(* IEC 61131-3 sources: plc-st-coding-agent/progress/evidence/f14_v10_full_20261113/jobs/custom_deepseek-v4pro (part 4) *)

(* ---- public-medium-02.raw_candidate_01.st ---- *)
TYPE ST_AnalogChannel :
STRUCT
    enable : BOOL;
    hiLIM : REAL;
    loLIM : REAL;
    bipolar : BOOL;
    measuringMode : INT;
    retVal : WORD;
    outputValue : REAL;
END_STRUCT
END_TYPE

(*
ENGINEERING_CONTRACT
Activation: process first count ordinal channels, count >= 0, clamped to min array lengths.
Enable: only channels[].enable = TRUE is evaluated; disabled rows retain previous retVal/outputValue.
retVal: for enabled rows write WORD#0 on success; WORD#16#8001 invalid measuringMode (PUB006); WORD#16#8002 hiLIM<=loLIM (PUB007).
Priority/simultaneous checks: measuringMode validity checked before hiLIM<=loLIM; simultaneous invalid mode and bad limits yields 16#8001 (unspecified, chosen).
outputValue: written only for enabled successful conversions; mode0 linear scaling clamped to 0/27648 or -27648/27648 (PUB003); mode1 raw/10 (PUB004); mode2 raw/100 (PUB005).
Read-only: analogValues unchanged; configuration fields only read (PUB001, PUB002).
Bounds: match by ordinal from each array lower bound; invalid count processes none.
Units: raw INT, output REAL, limits REAL; no time.
*)

(* CONTRACT_RULES [] *)

FUNCTION_BLOCK AnalogBatchProcessing
VAR_INPUT
    count : DINT;
END_VAR
VAR_IN_OUT
    analogValues : ARRAY[*] OF INT;
    channels : ARRAY[*] OF ST_AnalogChannel;
END_VAR
VAR
    tmp_lbA : DINT;
    tmp_lbC : DINT;
    tmp_availA : DINT;
    tmp_availC : DINT;
    tmp_process : DINT;
    tmp_i : DINT;
    tmp_idxA : DINT;
    tmp_idxC : DINT;
    tmp_raw : INT;
    tmp_rawReal : REAL;
    tmp_frac : REAL;
END_VAR

tmp_lbA := LOWER_BOUND(analogValues, 1);
tmp_lbC := LOWER_BOUND(channels, 1);
tmp_availA := UPPER_BOUND(analogValues, 1) - tmp_lbA + 1;
tmp_availC := UPPER_BOUND(channels, 1) - tmp_lbC + 1;

tmp_process := count;
IF tmp_process < 0 THEN
    tmp_process := 0;
END_IF;
IF tmp_process > tmp_availA THEN
    tmp_process := tmp_availA;
END_IF;
IF tmp_process > tmp_availC THEN
    tmp_process := tmp_availC;
END_IF;

FOR tmp_i := 0 TO tmp_process - 1 DO
    tmp_idxA := tmp_lbA + tmp_i;
    tmp_idxC := tmp_lbC + tmp_i;

    IF channels[tmp_idxC].enable THEN
        channels[tmp_idxC].retVal := WORD#0;

        IF (channels[tmp_idxC].measuringMode < 0) OR (channels[tmp_idxC].measuringMode > 2) THEN
            channels[tmp_idxC].retVal := WORD#16#8001;
            (* skip conversion; outputValue unchanged *)
        ELSIF channels[tmp_idxC].hiLIM <= channels[tmp_idxC].loLIM THEN
            channels[tmp_idxC].retVal := WORD#16#8002;
            (* skip conversion; outputValue unchanged *)
        ELSE
            tmp_raw := analogValues[tmp_idxA];
            tmp_rawReal := INT_TO_REAL(tmp_raw);

            CASE channels[tmp_idxC].measuringMode OF
                0:
                    IF channels[tmp_idxC].bipolar THEN
                        IF tmp_rawReal < -27648.0 THEN
                            tmp_rawReal := -27648.0;
                        ELSIF tmp_rawReal > 27648.0 THEN
                            tmp_rawReal := 27648.0;
                        END_IF;
                        tmp_frac := (tmp_rawReal + 27648.0) / 55296.0;
                    ELSE
                        IF tmp_rawReal < 0.0 THEN
                            tmp_rawReal := 0.0;
                        ELSIF tmp_rawReal > 27648.0 THEN
                            tmp_rawReal := 27648.0;
                        END_IF;
                        tmp_frac := tmp_rawReal / 27648.0;
                    END_IF;

                    channels[tmp_idxC].outputValue := channels[tmp_idxC].loLIM
                        + tmp_frac * (channels[tmp_idxC].hiLIM - channels[tmp_idxC].loLIM);

                1:
                    channels[tmp_idxC].outputValue := tmp_rawReal / 10.0;

                2:
                    channels[tmp_idxC].outputValue := tmp_rawReal / 100.0;

                ELSE
                    (* unreachable due to mode check above *)
                END_CASE;
        END_IF;
    END_IF;
END_FOR;

END_FUNCTION_BLOCK

(* ---- public-medium-02.raw_candidate_02.st ---- *)
TYPE ST_AnalogChannel :
STRUCT
    enable : BOOL;
    hiLIM : REAL;
    loLIM : REAL;
    bipolar : BOOL;
    measuringMode : INT;
    retVal : WORD;
    outputValue : REAL;
END_STRUCT
END_TYPE;

(*
ENGINEERING_CONTRACT
Activation: process first count ordinal channels, count >= 0, clamped to min array lengths.
Enable: only channels[].enable = TRUE is evaluated; disabled rows retain previous retVal/outputValue.
retVal: for enabled rows write WORD#0 on success; WORD#16#8001 invalid measuringMode (PUB006); WORD#16#8002 hiLIM<=loLIM (PUB007).
Priority/simultaneous checks: measuringMode validity checked before hiLIM<=loLIM; simultaneous invalid mode and bad limits yields 16#8001 (unspecified, chosen).
outputValue: written only for enabled successful conversions; mode0 linear scaling clamped to 0/27648 or -27648/27648 (PUB003); mode1 raw/10 (PUB004); mode2 raw/100 (PUB005).
Read-only: analogValues unchanged; configuration fields only read (PUB001, PUB002).
Bounds: match by ordinal from each array lower bound; invalid count processes none.
Units: raw INT, output REAL, limits REAL; no time.
*)

(* CONTRACT_RULES [] *)

FUNCTION_BLOCK AnalogBatchProcessing
VAR_INPUT
    count : DINT;
END_VAR
VAR_IN_OUT
    analogValues : ARRAY[*] OF INT;
    channels : ARRAY[*] OF ST_AnalogChannel;
END_VAR
VAR
    tmp_lbA : DINT;
    tmp_lbC : DINT;
    tmp_availA : DINT;
    tmp_availC : DINT;
    tmp_process : DINT;
    tmp_i : DINT;
    tmp_idxA : DINT;
    tmp_idxC : DINT;
    tmp_raw : INT;
    tmp_rawReal : REAL;
    tmp_frac : REAL;
END_VAR

tmp_lbA := LOWER_BOUND(analogValues, 1);
tmp_lbC := LOWER_BOUND(channels, 1);
tmp_availA := UPPER_BOUND(analogValues, 1) - tmp_lbA + 1;
tmp_availC := UPPER_BOUND(channels, 1) - tmp_lbC + 1;

tmp_process := count;
IF tmp_process < 0 THEN
    tmp_process := 0;
END_IF;
IF tmp_process > tmp_availA THEN
    tmp_process := tmp_availA;
END_IF;
IF tmp_process > tmp_availC THEN
    tmp_process := tmp_availC;
END_IF;

FOR tmp_i := 0 TO tmp_process - 1 DO
    tmp_idxA := tmp_lbA + tmp_i;
    tmp_idxC := tmp_lbC + tmp_i;

    IF channels[tmp_idxC].enable THEN
        channels[tmp_idxC].retVal := WORD#0;

        IF (channels[tmp_idxC].measuringMode < 0) OR (channels[tmp_idxC].measuringMode > 2) THEN
            channels[tmp_idxC].retVal := WORD#16#8001;
            (* skip conversion; outputValue unchanged *)
        ELSIF channels[tmp_idxC].hiLIM <= channels[tmp_idxC].loLIM THEN
            channels[tmp_idxC].retVal := WORD#16#8002;
            (* skip conversion; outputValue unchanged *)
        ELSE
            tmp_raw := analogValues[tmp_idxA];
            tmp_rawReal := INT_TO_REAL(tmp_raw);

            CASE channels[tmp_idxC].measuringMode OF
                0:
                    IF channels[tmp_idxC].bipolar THEN
                        IF tmp_rawReal < -27648.0 THEN
                            tmp_rawReal := -27648.0;
                        ELSIF tmp_rawReal > 27648.0 THEN
                            tmp_rawReal := 27648.0;
                        END_IF;
                        tmp_frac := (tmp_rawReal + 27648.0) / 55296.0;
                    ELSE
                        IF tmp_rawReal < 0.0 THEN
                            tmp_rawReal := 0.0;
                        ELSIF tmp_rawReal > 27648.0 THEN
                            tmp_rawReal := 27648.0;
                        END_IF;
                        tmp_frac := tmp_rawReal / 27648.0;
                    END_IF;

                    channels[tmp_idxC].outputValue := channels[tmp_idxC].loLIM
                        + tmp_frac * (channels[tmp_idxC].hiLIM - channels[tmp_idxC].loLIM);

                1:
                    channels[tmp_idxC].outputValue := tmp_rawReal / 10.0;

                2:
                    channels[tmp_idxC].outputValue := tmp_rawReal / 100.0;

                ELSE
                    (* unreachable due to mode check above *)
                    tmp_raw := tmp_raw;   (* dummy statement to satisfy CASE syntax *)
                END_CASE;
        END_IF;
    END_IF;
END_FOR;

END_FUNCTION_BLOCK

(* ---- public-medium-03.candidate_01.st ---- *)
FUNCTION_BLOCK FB
VAR_INPUT
    cyclicExecution : BOOL;
    trigger : BOOL;
    value : LREAL;
    windowSize : INT;
    reset : BOOL;
END_VAR
VAR_OUTPUT
    average : LREAL;
    windowSizeReached : BOOL;
    error : BOOL;
    status : WORD;
END_VAR
VAR
    local_triggerR : R_TRIG;
    local_buffer : ARRAY[0..99] OF LREAL;
    local_count : INT := 0;
    local_head : INT := 0;
    local_tail : INT := 0;
    local_sum : LREAL := 0.0;
END_VAR

(*
ENGINEERING_CONTRACT
average: update after accepted sample; holds between samples; reset clears to 0.0; invalid size preserves prior value (PUB001)
windowSizeReached: TRUE when buffered count >= windowSize; recalculated each valid scan; reset clears (PUB004)
error/status: invalid windowSize <1 or >100 sets error=TRUE status=16#8200; otherwise error=FALSE status=16#0000 (PUB003 PUB005 PUB006)
cyclicExecution: sample every scan; trigger has no effect while cyclicExecution=TRUE (PUB001)
trigger: sample on rising edge only when cyclicExecution=FALSE; edge detection runs every scan (PUB002)
reset: clears buffer/count/sum/average/windowSizeReached; then validates windowSize; reset scan does not sample (PUB003)
valid window size 1..100; circular buffer max 100; average = sum/count when count >0 else 0.0 (PUB005)
unspecified: valid windowSize change adapts by dropping oldest or appending to new size without automatic reset (PUB005)
*)
(* CONTRACT_RULES [] *)

BEGIN
    local_triggerR(CLK := trigger);

    IF reset THEN
        local_count := 0;
        local_head := 0;
        local_tail := 0;
        local_sum := 0.0;
        average := 0.0;
        windowSizeReached := FALSE;

        IF windowSize < 1 OR windowSize > 100 THEN
            error := TRUE;
            status := WORD#16#8200;
        ELSE
            error := FALSE;
            status := WORD#16#0000;
        END_IF;

        RETURN;
    END_IF;

    IF windowSize < 1 OR windowSize > 100 THEN
        error := TRUE;
        status := WORD#16#8200;
        windowSizeReached := FALSE;
        RETURN;
    ELSE
        error := FALSE;
        status := WORD#16#0000;
    END_IF;

    WHILE local_count > windowSize DO
        local_sum := local_sum - local_buffer[local_head];
        local_head := (local_head + 1) MOD 100;
        local_count := local_count - 1;
    END_WHILE;

    IF cyclicExecution OR local_triggerR.Q THEN
        IF local_count < windowSize THEN
            local_buffer[local_tail] := value;
            local_tail := (local_tail + 1) MOD 100;
            local_count := local_count + 1;
            local_sum := local_sum + value;
        ELSE
            local_sum := local_sum - local_buffer[local_head] + value;
            local_buffer[local_head] := value;
            local_head := (local_head + 1) MOD 100;
            local_tail := local_head;
        END_IF;
    END_IF;

    IF local_count > 0 THEN
        average := local_sum / INT_TO_LREAL(local_count);
    ELSE
        average := 0.0;
    END_IF;

    windowSizeReached := (local_count >= windowSize);
END_FUNCTION_BLOCK

(* ---- public-medium-03.candidate_02.st ---- *)
FUNCTION_BLOCK FB
VAR_INPUT
    cyclicExecution : BOOL;
    trigger : BOOL;
    value : LREAL;
    windowSize : INT;
    reset : BOOL;
END_VAR
VAR_OUTPUT
    average : LREAL;
    windowSizeReached : BOOL;
    error : BOOL;
    status : WORD;
END_VAR
VAR
    local_buffer : ARRAY[0..99] OF LREAL;
    local_count : INT := 0;
    local_head : INT := 0;
    local_tail : INT := 0;
    local_sum : LREAL := 0.0;
    local_trigger_prev : BOOL := FALSE;
    local_trigger_edge : BOOL := FALSE;
END_VAR

(*
ENGINEERING_CONTRACT
average: update after accepted sample; holds between samples; reset clears to 0.0; invalid size preserves prior value (PUB001)
windowSizeReached: TRUE when buffered count >= windowSize; recalculated each valid scan; reset clears (PUB004)
error/status: invalid windowSize <1 or >100 sets error=TRUE status=16#8200; otherwise error=FALSE status=16#0000 (PUB003 PUB005 PUB006)
cyclicExecution: sample every scan; trigger has no effect while cyclicExecution=TRUE (PUB001)
trigger: sample on rising edge only when cyclicExecution=FALSE; edge detection runs every scan (PUB002)
reset: clears buffer/count/sum/average/windowSizeReached; then validates windowSize; reset scan does not sample (PUB003)
valid window size 1..100; circular buffer max 100; average = sum/count when count >0 else 0.0 (PUB005)
unspecified: valid windowSize change adapts by dropping oldest or appending to new size without automatic reset (PUB005)
*)
(* CONTRACT_RULES [] *)

BEGIN
    local_trigger_edge := trigger AND NOT local_trigger_prev;
    local_trigger_prev := trigger;

    IF reset THEN
        local_count := 0;
        local_head := 0;
        local_tail := 0;
        local_sum := 0.0;
        average := 0.0;
        windowSizeReached := FALSE;

        IF windowSize < 1 OR windowSize > 100 THEN
            error := TRUE;
            status := WORD#16#8200;
        ELSE
            error := FALSE;
            status := WORD#16#0000;
        END_IF;

        RETURN;
    END_IF;

    IF windowSize < 1 OR windowSize > 100 THEN
        error := TRUE;
        status := WORD#16#8200;
        windowSizeReached := FALSE;
        RETURN;
    ELSE
        error := FALSE;
        status := WORD#16#0000;
    END_IF;

    WHILE local_count > windowSize DO
        local_sum := local_sum - local_buffer[local_head];
        local_head := (local_head + 1) MOD 100;
        local_count := local_count - 1;
    END_WHILE;

    IF cyclicExecution OR local_trigger_edge THEN
        IF local_count < windowSize THEN
            local_buffer[local_tail] := value;
            local_tail := (local_tail + 1) MOD 100;
            local_count := local_count + 1;
            local_sum := local_sum + value;
        ELSE
            local_sum := local_sum - local_buffer[local_head] + value;
            local_buffer[local_head] := value;
            local_head := (local_head + 1) MOD 100;
            local_tail := local_head;
        END_IF;
    END_IF;

    IF local_count > 0 THEN
        average := local_sum / INT_TO_LREAL(local_count);
    ELSE
        average := 0.0;
    END_IF;

    windowSizeReached := (local_count >= windowSize);
END_FUNCTION_BLOCK

(* ---- public-medium-03.candidate_03.st ---- *)
FUNCTION_BLOCK FB
VAR_INPUT
    cyclicExecution : BOOL;
    trigger : BOOL;
    value : LREAL;
    windowSize : INT;
    reset : BOOL;
END_VAR
VAR_OUTPUT
    average : LREAL;
    windowSizeReached : BOOL;
    error : BOOL;
    status : WORD;
END_VAR
VAR
    local_triggerPrev : BOOL;
    local_triggerRising : BOOL;
    local_buffer : ARRAY[0..99] OF LREAL;
    local_count : INT := 0;
    local_head : INT := 0;
    local_tail : INT := 0;
    local_sum : LREAL := 0.0;
END_VAR

(*
ENGINEERING_CONTRACT
average: update after accepted sample; holds between samples; reset clears to 0.0; invalid size preserves prior value (PUB001)
windowSizeReached: TRUE when buffered count >= windowSize; recalculated each valid scan; reset clears (PUB004)
error/status: invalid windowSize <1 or >100 sets error=TRUE status=16#8200; otherwise error=FALSE status=16#0000 (PUB003 PUB005 PUB006)
cyclicExecution: sample every scan; trigger has no effect while cyclicExecution=TRUE (PUB001)
trigger: sample on rising edge only when cyclicExecution=FALSE; edge detection runs every scan (PUB002)
reset: clears buffer/count/sum/average/windowSizeReached; then validates windowSize; reset scan does not sample (PUB003)
valid window size 1..100; circular buffer max 100; average = sum/count when count >0 else 0.0 (PUB005)
unspecified: valid windowSize change adapts by dropping oldest or appending to new size without automatic reset (PUB005)
*)
(* CONTRACT_RULES [] *)

BEGIN
    local_triggerRising := trigger AND NOT local_triggerPrev;
    local_triggerPrev := trigger;

    IF reset THEN
        local_count := 0;
        local_head := 0;
        local_tail := 0;
        local_sum := 0.0;
        average := 0.0;
        windowSizeReached := FALSE;

        IF windowSize < 1 OR windowSize > 100 THEN
            error := TRUE;
            status := WORD#16#8200;
        ELSE
            error := FALSE;
            status := WORD#16#0000;
        END_IF;

        RETURN;
    END_IF;

    IF windowSize < 1 OR windowSize > 100 THEN
        error := TRUE;
        status := WORD#16#8200;
        windowSizeReached := FALSE;
        RETURN;
    ELSE
        error := FALSE;
        status := WORD#16#0000;
    END_IF;

    WHILE local_count > windowSize DO
        local_sum := local_sum - local_buffer[local_head];
        local_head := (local_head + 1) MOD 100;
        local_count := local_count - 1;
    END_WHILE;

    IF cyclicExecution OR local_triggerRising THEN
        IF local_count < windowSize THEN
            local_buffer[local_tail] := value;
            local_tail := (local_tail + 1) MOD 100;
            local_count := local_count + 1;
            local_sum := local_sum + value;
        ELSE
            local_sum := local_sum - local_buffer[local_head] + value;
            local_buffer[local_head] := value;
            local_head := (local_head + 1) MOD 100;
            local_tail := (local_head + local_count) MOD 100;
        END_IF;
    END_IF;

    IF local_count > 0 THEN
        average := local_sum / INT_TO_LREAL(local_count);
    ELSE
        average := 0.0;
    END_IF;

    windowSizeReached := (local_count >= windowSize);
END_FUNCTION_BLOCK

(* ---- public-medium-03.candidate_04.st ---- *)
FUNCTION_BLOCK FB
VAR_INPUT
    cyclicExecution : BOOL;
    trigger : BOOL;
    value : LREAL;
    windowSize : INT;
    reset : BOOL;
END_VAR
VAR_OUTPUT
    average : LREAL;
    windowSizeReached : BOOL;
    error : BOOL;
    status : WORD;
END_VAR
VAR
    local_triggerR : R_TRIG;
    local_buffer : ARRAY[0..99] OF LREAL;
    local_count : INT := 0;
    local_head : INT := 0;
    local_tail : INT := 0;
    local_sum : LREAL := 0.0;
END_VAR

(*
ENGINEERING_CONTRACT
average: update after accepted sample; holds between samples; reset clears to 0.0; invalid size preserves prior value (PUB001)
windowSizeReached: TRUE when buffered count >= windowSize; recalculated each valid scan; reset clears (PUB004)
error/status: invalid windowSize <1 or >100 sets error=TRUE status=16#8200; otherwise error=FALSE status=16#0000 (PUB003 PUB005 PUB006)
cyclicExecution: sample every scan; trigger has no effect while cyclicExecution=TRUE (PUB001)
trigger: sample on rising edge only when cyclicExecution=FALSE; edge detection runs every scan (PUB002)
reset: clears buffer/count/sum/average/windowSizeReached; then validates windowSize; reset scan does not sample (PUB003)
valid window size 1..100; circular buffer max 100; average = sum/count when count >0 else 0.0 (PUB005)
unspecified: valid windowSize change adapts by dropping oldest or appending to new size without automatic reset (PUB005)
*)
(* CONTRACT_RULES [] *)

BEGIN
    local_triggerR(CLK := trigger);

    IF reset THEN
        local_count := 0;
        local_head := 0;
        local_tail := 0;
        local_sum := 0.0;
        average := 0.0;
        windowSizeReached := FALSE;

        IF windowSize < 1 OR windowSize > 100 THEN
            error := TRUE;
            status := WORD#16#8200;
        ELSE
            error := FALSE;
            status := WORD#16#0000;
        END_IF;

        RETURN;
    END_IF;

    IF windowSize < 1 OR windowSize > 100 THEN
        error := TRUE;
        status := WORD#16#8200;
        windowSizeReached := FALSE;
        RETURN;
    ELSE
        error := FALSE;
        status := WORD#16#0000;
    END_IF;

    WHILE local_count > windowSize DO
        local_sum := local_sum - local_buffer[local_head];
        local_head := (local_head + 1) MOD 100;
        local_count := local_count - 1;
    END_WHILE;

    IF cyclicExecution OR local_triggerR.Q THEN
        IF local_count < windowSize THEN
            local_buffer[local_tail] := value;
            local_tail := (local_tail + 1) MOD 100;
            local_count := local_count + 1;
            local_sum := local_sum + value;
        ELSE
            local_sum := local_sum - local_buffer[local_head] + value;
            local_buffer[local_head] := value;
            local_head := (local_head + 1) MOD 100;
            local_tail := local_head;
        END_IF;
    END_IF;

    IF local_count > 0 THEN
        average := local_sum / INT_TO_LREAL(local_count);
    ELSE
        average := 0.0;
    END_IF;

    windowSizeReached := (local_count >= windowSize);
END_FUNCTION_BLOCK

(* ---- public-medium-03.raw_candidate_01.st ---- *)
FUNCTION_BLOCK FB
VAR_INPUT
    cyclicExecution : BOOL;
    trigger : BOOL;
    value : LREAL;
    windowSize : INT;
    reset : BOOL;
END_VAR
VAR_OUTPUT
    average : LREAL;
    windowSizeReached : BOOL;
    error : BOOL;
    status : WORD;
END_VAR
VAR
    local_triggerR : R_TRIG;
    local_buffer : ARRAY[0..99] OF LREAL;
    local_count : INT := 0;
    local_head : INT := 0;
    local_tail : INT := 0;
    local_sum : LREAL := 0.0;
END_VAR

(*
ENGINEERING_CONTRACT
average: update after accepted sample; holds between samples; reset clears to 0.0; invalid size preserves prior value (PUB001)
windowSizeReached: TRUE when buffered count >= windowSize; recalculated each valid scan; reset clears (PUB004)
error/status: invalid windowSize <1 or >100 sets error=TRUE status=16#8200; otherwise error=FALSE status=16#0000 (PUB003 PUB005 PUB006)
cyclicExecution: sample every scan; trigger has no effect while cyclicExecution=TRUE (PUB001)
trigger: sample on rising edge only when cyclicExecution=FALSE; edge detection runs every scan (PUB002)
reset: clears buffer/count/sum/average/windowSizeReached; then validates windowSize; reset scan does not sample (PUB003)
valid window size 1..100; circular buffer max 100; average = sum/count when count >0 else 0.0 (PUB005)
unspecified: valid windowSize change adapts by dropping oldest or appending to new size without automatic reset (PUB005)
*)
(* CONTRACT_RULES [] *)

BEGIN
    local_triggerR(CLK := trigger);

    IF reset THEN
        local_count := 0;
        local_head := 0;
        local_tail := 0;
        local_sum := 0.0;
        average := 0.0;
        windowSizeReached := FALSE;

        IF windowSize < 1 OR windowSize > 100 THEN
            error := TRUE;
            status := WORD#16#8200;
        ELSE
            error := FALSE;
            status := WORD#16#0000;
        END_IF

        RETURN;
    END_IF

    IF windowSize < 1 OR windowSize > 100 THEN
        error := TRUE;
        status := WORD#16#8200;
        windowSizeReached := FALSE;
        RETURN;
    ELSE
        error := FALSE;
        status := WORD#16#0000;
    END_IF

    WHILE local_count > windowSize DO
        local_sum := local_sum - local_buffer[local_head];
        local_head := (local_head + 1) MOD 100;
        local_count := local_count - 1;
    END_WHILE

    IF cyclicExecution OR local_triggerR.Q THEN
        IF local_count < windowSize THEN
            local_buffer[local_tail] := value;
            local_tail := (local_tail + 1) MOD 100;
            local_count := local_count + 1;
            local_sum := local_sum + value;
        ELSE
            local_sum := local_sum - local_buffer[local_head] + value;
            local_buffer[local_head] := value;
            local_head := (local_head + 1) MOD 100;
            local_tail := local_head;
        END_IF
    END_IF

    IF local_count > 0 THEN
        average := local_sum / INT_TO_LREAL(local_count);
    ELSE
        average := 0.0;
    END_IF

    windowSizeReached := (local_count >= windowSize);
END_FUNCTION_BLOCK

(* ---- public-medium-03.raw_candidate_02.st ---- *)
FUNCTION_BLOCK FB
VAR_INPUT
    cyclicExecution : BOOL;
    trigger : BOOL;
    value : LREAL;
    windowSize : INT;
    reset : BOOL;
END_VAR
VAR_OUTPUT
    average : LREAL;
    windowSizeReached : BOOL;
    error : BOOL;
    status : WORD;
END_VAR
VAR
    local_buffer : ARRAY[0..99] OF LREAL;
    local_count : INT := 0;
    local_head : INT := 0;
    local_tail : INT := 0;
    local_sum : LREAL := 0.0;
    local_trigger_prev : BOOL := FALSE;
    local_trigger_edge : BOOL := FALSE;
END_VAR

(*
ENGINEERING_CONTRACT
average: update after accepted sample; holds between samples; reset clears to 0.0; invalid size preserves prior value (PUB001)
windowSizeReached: TRUE when buffered count >= windowSize; recalculated each valid scan; reset clears (PUB004)
error/status: invalid windowSize <1 or >100 sets error=TRUE status=16#8200; otherwise error=FALSE status=16#0000 (PUB003 PUB005 PUB006)
cyclicExecution: sample every scan; trigger has no effect while cyclicExecution=TRUE (PUB001)
trigger: sample on rising edge only when cyclicExecution=FALSE; edge detection runs every scan (PUB002)
reset: clears buffer/count/sum/average/windowSizeReached; then validates windowSize; reset scan does not sample (PUB003)
valid window size 1..100; circular buffer max 100; average = sum/count when count >0 else 0.0 (PUB005)
unspecified: valid windowSize change adapts by dropping oldest or appending to new size without automatic reset (PUB005)
*)
(* CONTRACT_RULES [] *)

BEGIN
    local_trigger_edge := trigger AND NOT local_trigger_prev;
    local_trigger_prev := trigger;

    IF reset THEN
        local_count := 0;
        local_head := 0;
        local_tail := 0;
        local_sum := 0.0;
        average := 0.0;
        windowSizeReached := FALSE;

        IF windowSize < 1 OR windowSize > 100 THEN
            error := TRUE;
            status := WORD#16#8200;
        ELSE
            error := FALSE;
            status := WORD#16#0000;
        END_IF;

        RETURN;
    END_IF;

    IF windowSize < 1 OR windowSize > 100 THEN
        error := TRUE;
        status := WORD#16#8200;
        windowSizeReached := FALSE;
        RETURN;
    ELSE
        error := FALSE;
        status := WORD#16#0000;
    END_IF;

    WHILE local_count > windowSize DO
        local_sum := local_sum - local_buffer[local_head];
        local_head := (local_head + 1) MOD 100;
        local_count := local_count - 1;
    END_WHILE;

    IF cyclicExecution OR local_trigger_edge THEN
        IF local_count < windowSize THEN
            local_buffer[local_tail] := value;
            local_tail := (local_tail + 1) MOD 100;
            local_count := local_count + 1;
            local_sum := local_sum + value;
        ELSE
            local_sum := local_sum - local_buffer[local_head] + value;
            local_buffer[local_head] := value;
            local_head := (local_head + 1) MOD 100;
            local_tail := local_head;
        END_IF;
    END_IF;

    IF local_count > 0 THEN
        average := local_sum / INT_TO_LREAL(local_count);
    ELSE
        average := 0.0;
    END_IF;

    windowSizeReached := (local_count >= windowSize);
END_FUNCTION_BLOCK

(* ---- public-medium-03.raw_candidate_03.st ---- *)
FUNCTION_BLOCK FB
VAR_INPUT
    cyclicExecution : BOOL;
    trigger : BOOL;
    value : LREAL;
    windowSize : INT;
    reset : BOOL;
END_VAR
VAR_OUTPUT
    average : LREAL;
    windowSizeReached : BOOL;
    error : BOOL;
    status : WORD;
END_VAR
VAR
    local_triggerPrev : BOOL;
    local_triggerRising : BOOL;
    local_buffer : ARRAY[0..99] OF LREAL;
    local_count : INT := 0;
    local_head : INT := 0;
    local_tail : INT := 0;
    local_sum : LREAL := 0.0;
END_VAR

(*
ENGINEERING_CONTRACT
average: update after accepted sample; holds between samples; reset clears to 0.0; invalid size preserves prior value (PUB001)
windowSizeReached: TRUE when buffered count >= windowSize; recalculated each valid scan; reset clears (PUB004)
error/status: invalid windowSize <1 or >100 sets error=TRUE status=16#8200; otherwise error=FALSE status=16#0000 (PUB003 PUB005 PUB006)
cyclicExecution: sample every scan; trigger has no effect while cyclicExecution=TRUE (PUB001)
trigger: sample on rising edge only when cyclicExecution=FALSE; edge detection runs every scan (PUB002)
reset: clears buffer/count/sum/average/windowSizeReached; then validates windowSize; reset scan does not sample (PUB003)
valid window size 1..100; circular buffer max 100; average = sum/count when count >0 else 0.0 (PUB005)
unspecified: valid windowSize change adapts by dropping oldest or appending to new size without automatic reset (PUB005)
*)
(* CONTRACT_RULES [] *)

BEGIN
    local_triggerRising := trigger AND NOT local_triggerPrev;
    local_triggerPrev := trigger;

    IF reset THEN
        local_count := 0;
        local_head := 0;
        local_tail := 0;
        local_sum := 0.0;
        average := 0.0;
        windowSizeReached := FALSE;

        IF windowSize < 1 OR windowSize > 100 THEN
            error := TRUE;
            status := WORD#16#8200;
        ELSE
            error := FALSE;
            status := WORD#16#0000;
        END_IF;

        RETURN;
    END_IF;

    IF windowSize < 1 OR windowSize > 100 THEN
        error := TRUE;
        status := WORD#16#8200;
        windowSizeReached := FALSE;
        RETURN;
    ELSE
        error := FALSE;
        status := WORD#16#0000;
    END_IF;

    WHILE local_count > windowSize DO
        local_sum := local_sum - local_buffer[local_head];
        local_head := (local_head + 1) MOD 100;
        local_count := local_count - 1;
    END_WHILE;

    IF cyclicExecution OR local_triggerRising THEN
        IF local_count < windowSize THEN
            local_buffer[local_tail] := value;
            local_tail := (local_tail + 1) MOD 100;
            local_count := local_count + 1;
            local_sum := local_sum + value;
        ELSE
            local_sum := local_sum - local_buffer[local_head] + value;
            local_buffer[local_head] := value;
            local_head := (local_head + 1) MOD 100;
            local_tail := (local_head + local_count) MOD 100;
        END_IF;
    END_IF;

    IF local_count > 0 THEN
        average := local_sum / INT_TO_LREAL(local_count);
    ELSE
        average := 0.0;
    END_IF;

    windowSizeReached := (local_count >= windowSize);
END_FUNCTION_BLOCK

(* ---- public-medium-03.raw_candidate_04.st ---- *)
FUNCTION_BLOCK FB
VAR_INPUT
    cyclicExecution : BOOL;
    trigger : BOOL;
    value : LREAL;
    windowSize : INT;
    reset : BOOL;
END_VAR
VAR_OUTPUT
    average : LREAL;
    windowSizeReached : BOOL;
    error : BOOL;
    status : WORD;
END_VAR
VAR
    local_triggerR : R_TRIG;
    local_buffer : ARRAY[0..99] OF LREAL;
    local_count : INT := 0;
    local_head : INT := 0;
    local_tail : INT := 0;
    local_sum : LREAL := 0.0;
END_VAR

(*
ENGINEERING_CONTRACT
average: update after accepted sample; holds between samples; reset clears to 0.0; invalid size preserves prior value (PUB001)
windowSizeReached: TRUE when buffered count >= windowSize; recalculated each valid scan; reset clears (PUB004)
error/status: invalid windowSize <1 or >100 sets error=TRUE status=16#8200; otherwise error=FALSE status=16#0000 (PUB003 PUB005 PUB006)
cyclicExecution: sample every scan; trigger has no effect while cyclicExecution=TRUE (PUB001)
trigger: sample on rising edge only when cyclicExecution=FALSE; edge detection runs every scan (PUB002)
reset: clears buffer/count/sum/average/windowSizeReached; then validates windowSize; reset scan does not sample (PUB003)
valid window size 1..100; circular buffer max 100; average = sum/count when count >0 else 0.0 (PUB005)
unspecified: valid windowSize change adapts by dropping oldest or appending to new size without automatic reset (PUB005)
*)
(* CONTRACT_RULES [] *)

BEGIN
    local_triggerR(CLK := trigger);

    IF reset THEN
        local_count := 0;
        local_head := 0;
        local_tail := 0;
        local_sum := 0.0;
        average := 0.0;
        windowSizeReached := FALSE;

        IF windowSize < 1 OR windowSize > 100 THEN
            error := TRUE;
            status := WORD#16#8200;
        ELSE
            error := FALSE;
            status := WORD#16#0000;
        END_IF;

        RETURN;
    END_IF;

    IF windowSize < 1 OR windowSize > 100 THEN
        error := TRUE;
        status := WORD#16#8200;
        windowSizeReached := FALSE;
        RETURN;
    ELSE
        error := FALSE;
        status := WORD#16#0000;
    END_IF;

    WHILE local_count > windowSize DO
        local_sum := local_sum - local_buffer[local_head];
        local_head := (local_head + 1) MOD 100;
        local_count := local_count - 1;
    END_WHILE;

    IF cyclicExecution OR local_triggerR.Q THEN
        IF local_count < windowSize THEN
            local_buffer[local_tail] := value;
            local_tail := (local_tail + 1) MOD 100;
            local_count := local_count + 1;
            local_sum := local_sum + value;
        ELSE
            local_sum := local_sum - local_buffer[local_head] + value;
            local_buffer[local_head] := value;
            local_head := (local_head + 1) MOD 100;
            local_tail := local_head;
        END_IF;
    END_IF;

    IF local_count > 0 THEN
        average := local_sum / INT_TO_LREAL(local_count);
    ELSE
        average := 0.0;
    END_IF;

    windowSizeReached := (local_count >= windowSize);
END_FUNCTION_BLOCK

(* ---- public-medium-04.candidate_01.st ---- *)
FUNCTION_BLOCK FB
VAR_INPUT
    TemperatureSensorInput : REAL;
    SetTemperature : REAL;
END_VAR
VAR_OUTPUT
    CurrentTemperature : REAL;
    SetTempDisplay : REAL;
    HeaterStatus : BOOL;
    OverheatProtection : BOOL;
    HeaterOutput : BOOL;
END_VAR
VAR
    tmp_heater_desired : BOOL := FALSE;
    local_heater_duration : TON;
    local_cooling_duration : TON;
    local_sensor_fault : BOOL;
END_VAR

(* ENGINEERING_CONTRACT
HeaterOutput: active <= sensor valid AND TemperatureSensorInput < SetTemperature (PUB003/PUB007).
OverheatProtection: latches when continuous HeaterOutput true >5s strict (T#5001MS); auto-lifts after 3s cooldown.
Fault: TemperatureSensorInput <0.0 or >100.0 forces heater off (PUB007).
Equal setpoint retains last heater command; initial off (unspecified).
Outputs reflect raw REAL/BOOL; HeaterStatus tracks HeaterOutput.
Same-scan priority: fault/overheat off over temp compare; overheat latch before output.
*)

(* CONTRACT_RULES [] *)

CurrentTemperature := TemperatureSensorInput;
SetTempDisplay := SetTemperature;

local_sensor_fault := (TemperatureSensorInput < 0.0) OR (TemperatureSensorInput > 100.0);

IF OverheatProtection THEN
    tmp_heater_desired := FALSE;
ELSE
    IF local_sensor_fault THEN
        tmp_heater_desired := FALSE;
    ELSE
        IF TemperatureSensorInput < SetTemperature THEN
            tmp_heater_desired := TRUE;
        ELSIF TemperatureSensorInput > SetTemperature THEN
            tmp_heater_desired := FALSE;
        END_IF;
    END_IF;
END_IF;

local_heater_duration(IN := tmp_heater_desired, PT := T#5001MS);

IF (NOT OverheatProtection) AND local_heater_duration.Q THEN
    OverheatProtection := TRUE;
    tmp_heater_desired := FALSE;
END_IF;

local_cooling_duration(IN := OverheatProtection, PT := T#3S);

IF OverheatProtection AND local_cooling_duration.Q THEN
    OverheatProtection := FALSE;
END_IF;

HeaterOutput := tmp_heater_desired;
HeaterStatus := HeaterOutput;

(* ---- public-medium-04.candidate_02.st ---- *)
FUNCTION_BLOCK FB
VAR_INPUT
    TemperatureSensorInput : REAL;
    SetTemperature : REAL;
END_VAR
VAR_OUTPUT
    CurrentTemperature : REAL;
    SetTempDisplay : REAL;
    HeaterStatus : BOOL;
    OverheatProtection : BOOL;
    HeaterOutput : BOOL;
END_VAR
VAR
    tmp_heater_desired : BOOL := FALSE;
    local_heater_duration : TON;
    local_cooling_duration : TON;
    local_sensor_fault : BOOL;
END_VAR

(* ENGINEERING_CONTRACT
HeaterOutput: active <= sensor valid AND TemperatureSensorInput < SetTemperature (PUB003/PUB007).
OverheatProtection: latches when continuous HeaterOutput true >5s strict (T#5001MS); auto-lifts after 3s cooldown.
Fault: TemperatureSensorInput <0.0 or >100.0 forces heater off (PUB007).
Equal setpoint retains last heater command; initial off (unspecified).
Outputs reflect raw REAL/BOOL; HeaterStatus tracks HeaterOutput.
Same-scan priority: fault/overheat off over temp compare; overheat latch before output.
*)

(* CONTRACT_RULES [] *)

CurrentTemperature := TemperatureSensorInput;
SetTempDisplay := SetTemperature;

local_sensor_fault := (TemperatureSensorInput < 0.0) OR (TemperatureSensorInput > 100.0);

IF OverheatProtection THEN
    tmp_heater_desired := FALSE;
ELSE
    IF local_sensor_fault THEN
        tmp_heater_desired := FALSE;
    ELSE
        IF TemperatureSensorInput < SetTemperature THEN
            tmp_heater_desired := TRUE;
        ELSIF TemperatureSensorInput > SetTemperature THEN
            tmp_heater_desired := FALSE;
        END_IF;
    END_IF;
END_IF;

local_heater_duration(IN := tmp_heater_desired, PT := T#5001MS);

IF (NOT OverheatProtection) AND local_heater_duration.Q THEN
    OverheatProtection := TRUE;
    tmp_heater_desired := FALSE;
END_IF;

local_cooling_duration(IN := OverheatProtection, PT := T#3S);

IF OverheatProtection AND local_cooling_duration.Q THEN
    OverheatProtection := FALSE;
END_IF;

HeaterOutput := tmp_heater_desired;
HeaterStatus := HeaterOutput;

END_FUNCTION_BLOCK

(* ---- public-medium-04.candidate_03.st ---- *)
FUNCTION_BLOCK FB
VAR_INPUT
    TemperatureSensorInput : REAL;
    SetTemperature : REAL;
END_VAR
VAR_OUTPUT
    CurrentTemperature : REAL;
    SetTempDisplay : REAL;
    HeaterStatus : BOOL;
    OverheatProtection : BOOL;
    HeaterOutput : BOOL;
END_VAR
VAR
    tmp_heater_desired : BOOL := FALSE;
    local_heater_duration : TON;
    local_cooling_duration : TON;
    local_sensor_fault : BOOL;
    local_heater_request : BOOL := FALSE;
END_VAR

(* ENGINEERING_CONTRACT
HeaterOutput: active <= sensor valid AND TemperatureSensorInput < SetTemperature, unless OverheatProtection active (PUB003/PUB004/PUB007).
OverheatProtection: latches when continuous HeaterOutput true >5s strict (T#5001MS); auto-lifts after 3s cooldown (T#3S).
Fault: TemperatureSensorInput <0.0 or >100.0 forces heater off (PUB007).
Equal setpoint retains last heater request; initial request off (unspecified).
Outputs reflect raw REAL/BOOL; HeaterStatus tracks HeaterOutput.
Same-scan priority: fault/overheat off over temp compare; cooldown reset immediately restores heater request.
*)

(* CONTRACT_RULES [] *)

CurrentTemperature := TemperatureSensorInput;
SetTempDisplay := SetTemperature;

local_sensor_fault := (TemperatureSensorInput < 0.0) OR (TemperatureSensorInput > 100.0);

IF local_sensor_fault THEN
    local_heater_request := FALSE;
ELSE
    IF TemperatureSensorInput < SetTemperature THEN
        local_heater_request := TRUE;
    ELSIF TemperatureSensorInput > SetTemperature THEN
        local_heater_request := FALSE;
    END_IF;
END_IF;

tmp_heater_desired := local_heater_request AND NOT OverheatProtection;

local_heater_duration(IN := tmp_heater_desired, PT := T#5001MS);

IF (NOT OverheatProtection) AND local_heater_duration.Q THEN
    OverheatProtection := TRUE;
    tmp_heater_desired := FALSE;
END_IF;

local_cooling_duration(IN := OverheatProtection, PT := T#3S);

IF OverheatProtection AND local_cooling_duration.Q THEN
    OverheatProtection := FALSE;
    tmp_heater_desired := local_heater_request AND NOT OverheatProtection;
    local_heater_duration(IN := tmp_heater_desired, PT := T#5001MS);
END_IF;

HeaterOutput := tmp_heater_desired;
HeaterStatus := HeaterOutput;

END_FUNCTION_BLOCK

(* ---- public-medium-04.raw_candidate_01.st ---- *)
FUNCTION_BLOCK FB
VAR_INPUT
    TemperatureSensorInput : REAL;
    SetTemperature : REAL;
END_VAR
VAR_OUTPUT
    CurrentTemperature : REAL;
    SetTempDisplay : REAL;
    HeaterStatus : BOOL;
    OverheatProtection : BOOL;
    HeaterOutput : BOOL;
END_VAR
VAR
    tmp_heater_desired : BOOL := FALSE;
    local_heater_duration : TON;
    local_cooling_duration : TON;
    local_sensor_fault : BOOL;
END_VAR

(* ENGINEERING_CONTRACT
HeaterOutput: active <= sensor valid AND TemperatureSensorInput < SetTemperature (PUB003/PUB007).
OverheatProtection: latches when continuous HeaterOutput true >5s strict (T#5001MS); auto-lifts after 3s cooldown.
Fault: TemperatureSensorInput <0.0 or >100.0 forces heater off (PUB007).
Equal setpoint retains last heater command; initial off (unspecified).
Outputs reflect raw REAL/BOOL; HeaterStatus tracks HeaterOutput.
Same-scan priority: fault/overheat off over temp compare; overheat latch before output.
*)

(* CONTRACT_RULES [] *)

CurrentTemperature := TemperatureSensorInput;
SetTempDisplay := SetTemperature;

local_sensor_fault := (TemperatureSensorInput < 0.0) OR (TemperatureSensorInput > 100.0);

IF OverheatProtection THEN
    tmp_heater_desired := FALSE;
ELSE
    IF local_sensor_fault THEN
        tmp_heater_desired := FALSE;
    ELSE
        IF TemperatureSensorInput < SetTemperature THEN
            tmp_heater_desired := TRUE;
        ELSIF TemperatureSensorInput > SetTemperature THEN
            tmp_heater_desired := FALSE;
        END_IF;
    END_IF;
END_IF;

local_heater_duration(IN := tmp_heater_desired, PT := T#5001MS);

IF (NOT OverheatProtection) AND local_heater_duration.Q THEN
    OverheatProtection := TRUE;
    tmp_heater_desired := FALSE;
END_IF;

local_cooling_duration(IN := OverheatProtection, PT := T#3S);

IF OverheatProtection AND local_cooling_duration.Q THEN
    OverheatProtection := FALSE;
END_IF;

HeaterOutput := tmp_heater_desired;
HeaterStatus := HeaterOutput;

(* ---- public-medium-04.raw_candidate_02.st ---- *)
FUNCTION_BLOCK FB
VAR_INPUT
    TemperatureSensorInput : REAL;
    SetTemperature : REAL;
END_VAR
VAR_OUTPUT
    CurrentTemperature : REAL;
    SetTempDisplay : REAL;
    HeaterStatus : BOOL;
    OverheatProtection : BOOL;
    HeaterOutput : BOOL;
END_VAR
VAR
    tmp_heater_desired : BOOL := FALSE;
    local_heater_duration : TON;
    local_cooling_duration : TON;
    local_sensor_fault : BOOL;
END_VAR

(* ENGINEERING_CONTRACT
HeaterOutput: active <= sensor valid AND TemperatureSensorInput < SetTemperature (PUB003/PUB007).
OverheatProtection: latches when continuous HeaterOutput true >5s strict (T#5001MS); auto-lifts after 3s cooldown.
Fault: TemperatureSensorInput <0.0 or >100.0 forces heater off (PUB007).
Equal setpoint retains last heater command; initial off (unspecified).
Outputs reflect raw REAL/BOOL; HeaterStatus tracks HeaterOutput.
Same-scan priority: fault/overheat off over temp compare; overheat latch before output.
*)

(* CONTRACT_RULES [] *)

CurrentTemperature := TemperatureSensorInput;
SetTempDisplay := SetTemperature;

local_sensor_fault := (TemperatureSensorInput < 0.0) OR (TemperatureSensorInput > 100.0);

IF OverheatProtection THEN
    tmp_heater_desired := FALSE;
ELSE
    IF local_sensor_fault THEN
        tmp_heater_desired := FALSE;
    ELSE
        IF TemperatureSensorInput < SetTemperature THEN
            tmp_heater_desired := TRUE;
        ELSIF TemperatureSensorInput > SetTemperature THEN
            tmp_heater_desired := FALSE;
        END_IF;
    END_IF;
END_IF;

local_heater_duration(IN := tmp_heater_desired, PT := T#5001MS);

IF (NOT OverheatProtection) AND local_heater_duration.Q THEN
    OverheatProtection := TRUE;
    tmp_heater_desired := FALSE;
END_IF;

local_cooling_duration(IN := OverheatProtection, PT := T#3S);

IF OverheatProtection AND local_cooling_duration.Q THEN
    OverheatProtection := FALSE;
END_IF;

HeaterOutput := tmp_heater_desired;
HeaterStatus := HeaterOutput;

END_FUNCTION_BLOCK

(* ---- public-medium-04.raw_candidate_03.st ---- *)
FUNCTION_BLOCK FB
VAR_INPUT
    TemperatureSensorInput : REAL;
    SetTemperature : REAL;
END_VAR
VAR_OUTPUT
    CurrentTemperature : REAL;
    SetTempDisplay : REAL;
    HeaterStatus : BOOL;
    OverheatProtection : BOOL;
    HeaterOutput : BOOL;
END_VAR
VAR
    tmp_heater_desired : BOOL := FALSE;
    local_heater_duration : TON;
    local_cooling_duration : TON;
    local_sensor_fault : BOOL;
    local_heater_request : BOOL := FALSE;
END_VAR

(* ENGINEERING_CONTRACT
HeaterOutput: active <= sensor valid AND TemperatureSensorInput < SetTemperature, unless OverheatProtection active (PUB003/PUB004/PUB007).
OverheatProtection: latches when continuous HeaterOutput true >5s strict (T#5001MS); auto-lifts after 3s cooldown (T#3S).
Fault: TemperatureSensorInput <0.0 or >100.0 forces heater off (PUB007).
Equal setpoint retains last heater request; initial request off (unspecified).
Outputs reflect raw REAL/BOOL; HeaterStatus tracks HeaterOutput.
Same-scan priority: fault/overheat off over temp compare; cooldown reset immediately restores heater request.
*)

(* CONTRACT_RULES [] *)

CurrentTemperature := TemperatureSensorInput;
SetTempDisplay := SetTemperature;

local_sensor_fault := (TemperatureSensorInput < 0.0) OR (TemperatureSensorInput > 100.0);

IF local_sensor_fault THEN
    local_heater_request := FALSE;
ELSE
    IF TemperatureSensorInput < SetTemperature THEN
        local_heater_request := TRUE;
    ELSIF TemperatureSensorInput > SetTemperature THEN
        local_heater_request := FALSE;
    END_IF;
END_IF;

tmp_heater_desired := local_heater_request AND NOT OverheatProtection;

local_heater_duration(IN := tmp_heater_desired, PT := T#5001MS);

IF (NOT OverheatProtection) AND local_heater_duration.Q THEN
    OverheatProtection := TRUE;
    tmp_heater_desired := FALSE;
END_IF;

local_cooling_duration(IN := OverheatProtection, PT := T#3S);

IF OverheatProtection AND local_cooling_duration.Q THEN
    OverheatProtection := FALSE;
    tmp_heater_desired := local_heater_request AND NOT OverheatProtection;
    local_heater_duration(IN := tmp_heater_desired, PT := T#5001MS);
END_IF;

HeaterOutput := tmp_heater_desired;
HeaterStatus := HeaterOutput;

END_FUNCTION_BLOCK

(* ---- public-medium-05.candidate_01.st ---- *)
FUNCTION_BLOCK ProductionLineControl
VAR
    trigA : R_TRIG;
    trigB : R_TRIG;
    trigC : R_TRIG;
    movingToB : BOOL := FALSE;
    movingToC : BOOL := FALSE;
    completionLatched : BOOL := FALSE;
END_VAR

(* ENGINEERING_CONTRACT
MotorForward: manual = ForwardButton AND NOT ReverseButton;
  auto = movingToB OR movingToC. Hold until target sensor or mode change.
MotorReverse: manual = ReverseButton AND NOT ForwardButton;
  interlocked, both buttons => neither. No auto reverse.
CompletionLight: auto only, set on ButtonC rising edge while SensorC true,
  reset when SensorC false or mode manual. Unspecified manual completion light = off.
State movingToB/movingToC: start on source button rising edge at source sensor,
  stop on target sensor. Cleared in manual.
State completionLatched: holds until SensorC false or mode manual.
PUB001-PUB008 satisfied.
*)
(* CONTRACT_RULES [] *)

trigA(CLK := ButtonA);
trigB(CLK := ButtonB);
trigC(CLK := ButtonC);

MotorForward := FALSE;
MotorReverse := FALSE;
CompletionLight := FALSE;

IF Mode THEN
    (* Automatic mode *)
    MotorReverse := FALSE;

    (* Arrival stops first: product reached target station *)
    IF movingToB AND SensorB THEN
        movingToB := FALSE;
    END_IF;

    IF movingToC AND SensorC THEN
        movingToC := FALSE;
    END_IF;

    (* Start movement or completion when not already moving *)
    IF NOT movingToB AND NOT movingToC THEN
        IF SensorA AND trigA.Q THEN
            movingToB := TRUE;
        ELSIF SensorB AND trigB.Q THEN
            movingToC := TRUE;
        ELSIF SensorC AND trigC.Q THEN
            completionLatched := TRUE;
        END_IF;
    END_IF;

    (* Completion light off when product is taken away from C *)
    IF NOT SensorC THEN
        completionLatched := FALSE;
    END_IF;

    CompletionLight := completionLatched;
    MotorForward := movingToB OR movingToC;
ELSE
    (* Manual mode: clear all automatic sequence state *)
    movingToB := FALSE;
    movingToC := FALSE;
    completionLatched := FALSE;

    IF ForwardButton AND NOT ReverseButton THEN
        MotorForward := TRUE;
        MotorReverse := FALSE;
    ELSIF ReverseButton AND NOT ForwardButton THEN
        MotorForward := FALSE;
        MotorReverse := TRUE;
    ELSE
        MotorForward := FALSE;
        MotorReverse := FALSE;
    END_IF;

    CompletionLight := FALSE;
END_IF;
END_FUNCTION_BLOCK

(* ---- public-medium-05.candidate_02.st ---- *)
FUNCTION_BLOCK ProductionLineControl
VAR_INPUT
    Mode : BOOL;
    ForwardButton : BOOL;
    ReverseButton : BOOL;
    SensorA : BOOL;
    SensorB : BOOL;
    SensorC : BOOL;
    ButtonA : BOOL;
    ButtonB : BOOL;
    ButtonC : BOOL;
END_VAR
VAR_OUTPUT
    MotorForward : BOOL;
    MotorReverse : BOOL;
    CompletionLight : BOOL;
END_VAR
VAR
    trigA : R_TRIG;
    trigB : R_TRIG;
    trigC : R_TRIG;
    movingToB : BOOL := FALSE;
    movingToC : BOOL := FALSE;
    completionLatched : BOOL := FALSE;
END_VAR

(* ENGINEERING_CONTRACT
MotorForward: manual = ForwardButton AND NOT ReverseButton;
  auto = movingToB OR movingToC. Hold until target sensor or mode change.
MotorReverse: manual = ReverseButton AND NOT ForwardButton;
  interlocked, both buttons => neither. No auto reverse.
CompletionLight: auto only, set on ButtonC rising edge while SensorC true,
  reset when SensorC false or mode manual. Unspecified manual completion light = off.
State movingToB/movingToC: start on source button rising edge at source sensor,
  stop on target sensor. Cleared in manual.
State completionLatched: holds until SensorC false or mode manual.
PUB001-PUB008 satisfied.
*)
(* CONTRACT_RULES [] *)

trigA(CLK := ButtonA);
trigB(CLK := ButtonB);
trigC(CLK := ButtonC);

MotorForward := FALSE;
MotorReverse := FALSE;
CompletionLight := FALSE;

IF Mode THEN
    (* Automatic mode *)
    MotorReverse := FALSE;

    (* Arrival stops first: product reached target station *)
    IF movingToB AND SensorB THEN
        movingToB := FALSE;
    END_IF;

    IF movingToC AND SensorC THEN
        movingToC := FALSE;
    END_IF;

    (* Start movement or completion when not already moving *)
    IF NOT movingToB AND NOT movingToC THEN
        IF SensorA AND trigA.Q THEN
            movingToB := TRUE;
        ELSIF SensorB AND trigB.Q THEN
            movingToC := TRUE;
        ELSIF SensorC AND trigC.Q THEN
            completionLatched := TRUE;
        END_IF;
    END_IF;

    (* Completion light off when product is taken away from C *)
    IF NOT SensorC THEN
        completionLatched := FALSE;
    END_IF;

    CompletionLight := completionLatched;
    MotorForward := movingToB OR movingToC;
ELSE
    (* Manual mode: clear all automatic sequence state *)
    movingToB := FALSE;
    movingToC := FALSE;
    completionLatched := FALSE;

    IF ForwardButton AND NOT ReverseButton THEN
        MotorForward := TRUE;
        MotorReverse := FALSE;
    ELSIF ReverseButton AND NOT ForwardButton THEN
        MotorForward := FALSE;
        MotorReverse := TRUE;
    ELSE
        MotorForward := FALSE;
        MotorReverse := FALSE;
    END_IF;

    CompletionLight := FALSE;
END_IF;
END_FUNCTION_BLOCK

(* ---- public-medium-05.candidate_03.st ---- *)
FUNCTION_BLOCK ProductionLineControl
VAR_INPUT
    Mode : BOOL;
    ForwardButton : BOOL;
    ReverseButton : BOOL;
    SensorA : BOOL;
    SensorB : BOOL;
    SensorC : BOOL;
    ButtonA : BOOL;
    ButtonB : BOOL;
    ButtonC : BOOL;
END_VAR
VAR_OUTPUT
    MotorForward : BOOL;
    MotorReverse : BOOL;
    CompletionLight : BOOL;
END_VAR
VAR
    movingToB : BOOL := FALSE;
    movingToC : BOOL := FALSE;
    completionLatched : BOOL := FALSE;
END_VAR

(* ENGINEERING_CONTRACT
MotorForward: manual = ForwardButton AND NOT ReverseButton;
  auto = movingToB OR movingToC. Hold until target sensor or mode change.
MotorReverse: manual = ReverseButton AND NOT ForwardButton;
  interlocked, both buttons => neither. No auto reverse.
CompletionLight: auto only, set when SensorC AND ButtonC true (level),
  reset when SensorC false or mode manual. Unspecified manual completion light = off.
State movingToB/movingToC: start when source sensor AND corresponding button true,
  stop on target sensor. Cleared in manual.
State completionLatched: holds until SensorC false or mode manual.
All automatic actions level-triggered (button held is sufficient) per public wording.
PUB001-PUB008 satisfied.
*)
(* CONTRACT_RULES [] *)

MotorForward := FALSE;
MotorReverse := FALSE;
CompletionLight := FALSE;

IF Mode THEN
    (* Automatic mode *)
    MotorReverse := FALSE;

    (* Arrival stops first: product reached target station *)
    IF movingToB AND SensorB THEN
        movingToB := FALSE;
    END_IF;

    IF movingToC AND SensorC THEN
        movingToC := FALSE;
    END_IF;

    (* Start movement or completion when not already moving *)
    IF NOT movingToB AND NOT movingToC THEN
        IF SensorA AND ButtonA THEN
            movingToB := TRUE;
        ELSIF SensorB AND ButtonB THEN
            movingToC := TRUE;
        ELSIF SensorC AND ButtonC THEN
            completionLatched := TRUE;
        END_IF;
    END_IF;

    (* Completion light off when product is taken away from C *)
    IF NOT SensorC THEN
        completionLatched := FALSE;
    END_IF;

    CompletionLight := completionLatched;
    MotorForward := movingToB OR movingToC;
ELSE
    (* Manual mode: clear all automatic sequence state *)
    movingToB := FALSE;
    movingToC := FALSE;
    completionLatched := FALSE;

    IF ForwardButton AND NOT ReverseButton THEN
        MotorForward := TRUE;
        MotorReverse := FALSE;
    ELSIF ReverseButton AND NOT ForwardButton THEN
        MotorForward := FALSE;
        MotorReverse := TRUE;
    ELSE
        MotorForward := FALSE;
        MotorReverse := FALSE;
    END_IF;

    CompletionLight := FALSE;
END_IF;
END_FUNCTION_BLOCK

(* ---- public-medium-05.raw_candidate_01.st ---- *)
FUNCTION_BLOCK ProductionLineControl
VAR
    trigA : R_TRIG;
    trigB : R_TRIG;
    trigC : R_TRIG;
    movingToB : BOOL := FALSE;
    movingToC : BOOL := FALSE;
    completionLatched : BOOL := FALSE;
END_VAR

(* ENGINEERING_CONTRACT
MotorForward: manual = ForwardButton AND NOT ReverseButton;
  auto = movingToB OR movingToC. Hold until target sensor or mode change.
MotorReverse: manual = ReverseButton AND NOT ForwardButton;
  interlocked, both buttons => neither. No auto reverse.
CompletionLight: auto only, set on ButtonC rising edge while SensorC true,
  reset when SensorC false or mode manual. Unspecified manual completion light = off.
State movingToB/movingToC: start on source button rising edge at source sensor,
  stop on target sensor. Cleared in manual.
State completionLatched: holds until SensorC false or mode manual.
PUB001-PUB008 satisfied.
*)
(* CONTRACT_RULES [] *)

trigA(CLK := ButtonA);
trigB(CLK := ButtonB);
trigC(CLK := ButtonC);

MotorForward := FALSE;
MotorReverse := FALSE;
CompletionLight := FALSE;

IF Mode THEN
    (* Automatic mode *)
    MotorReverse := FALSE;

    (* Arrival stops first: product reached target station *)
    IF movingToB AND SensorB THEN
        movingToB := FALSE;
    END_IF;

    IF movingToC AND SensorC THEN
        movingToC := FALSE;
    END_IF;

    (* Start movement or completion when not already moving *)
    IF NOT movingToB AND NOT movingToC THEN
        IF SensorA AND trigA.Q THEN
            movingToB := TRUE;
        ELSIF SensorB AND trigB.Q THEN
            movingToC := TRUE;
        ELSIF SensorC AND trigC.Q THEN
            completionLatched := TRUE;
        END_IF;
    END_IF;

    (* Completion light off when product is taken away from C *)
    IF NOT SensorC THEN
        completionLatched := FALSE;
    END_IF;

    CompletionLight := completionLatched;
    MotorForward := movingToB OR movingToC;
ELSE
    (* Manual mode: clear all automatic sequence state *)
    movingToB := FALSE;
    movingToC := FALSE;
    completionLatched := FALSE;

    IF ForwardButton AND NOT ReverseButton THEN
        MotorForward := TRUE;
        MotorReverse := FALSE;
    ELSIF ReverseButton AND NOT ForwardButton THEN
        MotorForward := FALSE;
        MotorReverse := TRUE;
    ELSE
        MotorForward := FALSE;
        MotorReverse := FALSE;
    END_IF;

    CompletionLight := FALSE;
END_IF;
END_FUNCTION_BLOCK

(* ---- public-medium-05.raw_candidate_02.st ---- *)
FUNCTION_BLOCK ProductionLineControl
VAR_INPUT
    Mode : BOOL;
    ForwardButton : BOOL;
    ReverseButton : BOOL;
    SensorA : BOOL;
    SensorB : BOOL;
    SensorC : BOOL;
    ButtonA : BOOL;
    ButtonB : BOOL;
    ButtonC : BOOL;
END_VAR
VAR_OUTPUT
    MotorForward : BOOL;
    MotorReverse : BOOL;
    CompletionLight : BOOL;
END_VAR
VAR
    trigA : R_TRIG;
    trigB : R_TRIG;
    trigC : R_TRIG;
    movingToB : BOOL := FALSE;
    movingToC : BOOL := FALSE;
    completionLatched : BOOL := FALSE;
END_VAR

(* ENGINEERING_CONTRACT
MotorForward: manual = ForwardButton AND NOT ReverseButton;
  auto = movingToB OR movingToC. Hold until target sensor or mode change.
MotorReverse: manual = ReverseButton AND NOT ForwardButton;
  interlocked, both buttons => neither. No auto reverse.
CompletionLight: auto only, set on ButtonC rising edge while SensorC true,
  reset when SensorC false or mode manual. Unspecified manual completion light = off.
State movingToB/movingToC: start on source button rising edge at source sensor,
  stop on target sensor. Cleared in manual.
State completionLatched: holds until SensorC false or mode manual.
PUB001-PUB008 satisfied.
*)
(* CONTRACT_RULES [] *)

trigA(CLK := ButtonA);
trigB(CLK := ButtonB);
trigC(CLK := ButtonC);

MotorForward := FALSE;
MotorReverse := FALSE;
CompletionLight := FALSE;

IF Mode THEN
    (* Automatic mode *)
    MotorReverse := FALSE;

    (* Arrival stops first: product reached target station *)
    IF movingToB AND SensorB THEN
        movingToB := FALSE;
    END_IF;

    IF movingToC AND SensorC THEN
        movingToC := FALSE;
    END_IF;

    (* Start movement or completion when not already moving *)
    IF NOT movingToB AND NOT movingToC THEN
        IF SensorA AND trigA.Q THEN
            movingToB := TRUE;
        ELSIF SensorB AND trigB.Q THEN
            movingToC := TRUE;
        ELSIF SensorC AND trigC.Q THEN
            completionLatched := TRUE;
        END_IF;
    END_IF;

    (* Completion light off when product is taken away from C *)
    IF NOT SensorC THEN
        completionLatched := FALSE;
    END_IF;

    CompletionLight := completionLatched;
    MotorForward := movingToB OR movingToC;
ELSE
    (* Manual mode: clear all automatic sequence state *)
    movingToB := FALSE;
    movingToC := FALSE;
    completionLatched := FALSE;

    IF ForwardButton AND NOT ReverseButton THEN
        MotorForward := TRUE;
        MotorReverse := FALSE;
    ELSIF ReverseButton AND NOT ForwardButton THEN
        MotorForward := FALSE;
        MotorReverse := TRUE;
    ELSE
        MotorForward := FALSE;
        MotorReverse := FALSE;
    END_IF;

    CompletionLight := FALSE;
END_IF;
END_FUNCTION_BLOCK

(* ---- public-medium-05.raw_candidate_03.st ---- *)
FUNCTION_BLOCK ProductionLineControl
VAR_INPUT
    Mode : BOOL;
    ForwardButton : BOOL;
    ReverseButton : BOOL;
    SensorA : BOOL;
    SensorB : BOOL;
    SensorC : BOOL;
    ButtonA : BOOL;
    ButtonB : BOOL;
    ButtonC : BOOL;
END_VAR
VAR_OUTPUT
    MotorForward : BOOL;
    MotorReverse : BOOL;
    CompletionLight : BOOL;
END_VAR
VAR
    movingToB : BOOL := FALSE;
    movingToC : BOOL := FALSE;
    completionLatched : BOOL := FALSE;
END_VAR

(* ENGINEERING_CONTRACT
MotorForward: manual = ForwardButton AND NOT ReverseButton;
  auto = movingToB OR movingToC. Hold until target sensor or mode change.
MotorReverse: manual = ReverseButton AND NOT ForwardButton;
  interlocked, both buttons => neither. No auto reverse.
CompletionLight: auto only, set when SensorC AND ButtonC true (level),
  reset when SensorC false or mode manual. Unspecified manual completion light = off.
State movingToB/movingToC: start when source sensor AND corresponding button true,
  stop on target sensor. Cleared in manual.
State completionLatched: holds until SensorC false or mode manual.
All automatic actions level-triggered (button held is sufficient) per public wording.
PUB001-PUB008 satisfied.
*)
(* CONTRACT_RULES [] *)

MotorForward := FALSE;
MotorReverse := FALSE;
CompletionLight := FALSE;

IF Mode THEN
    (* Automatic mode *)
    MotorReverse := FALSE;

    (* Arrival stops first: product reached target station *)
    IF movingToB AND SensorB THEN
        movingToB := FALSE;
    END_IF;

    IF movingToC AND SensorC THEN
        movingToC := FALSE;
    END_IF;

    (* Start movement or completion when not already moving *)
    IF NOT movingToB AND NOT movingToC THEN
        IF SensorA AND ButtonA THEN
            movingToB := TRUE;
        ELSIF SensorB AND ButtonB THEN
            movingToC := TRUE;
        ELSIF SensorC AND ButtonC THEN
            completionLatched := TRUE;
        END_IF;
    END_IF;

    (* Completion light off when product is taken away from C *)
    IF NOT SensorC THEN
        completionLatched := FALSE;
    END_IF;

    CompletionLight := completionLatched;
    MotorForward := movingToB OR movingToC;
ELSE
    (* Manual mode: clear all automatic sequence state *)
    movingToB := FALSE;
    movingToC := FALSE;
    completionLatched := FALSE;

    IF ForwardButton AND NOT ReverseButton THEN
        MotorForward := TRUE;
        MotorReverse := FALSE;
    ELSIF ReverseButton AND NOT ForwardButton THEN
        MotorForward := FALSE;
        MotorReverse := TRUE;
    ELSE
        MotorForward := FALSE;
        MotorReverse := FALSE;
    END_IF;

    CompletionLight := FALSE;
END_IF;
END_FUNCTION_BLOCK

(* ---- public-medium-06.candidate_01.st ---- *)
FUNCTION_BLOCK SlabThicknessFaultMonitor
VAR_INPUT
    THICKNESS_FAULT : BOOL;
    THICKNESS_SIGNAL_VALID : BOOL;
    CUTTING_RUN : BOOL;
    FaultTimestamp : DINT;
    CycleTime : TIME;
END_VAR
VAR_OUTPUT
    THICKNESS_ALARM : BOOL;
    Slab_Fault_Counter : UINT;
    Slab_Runtime_Accumulator : LTIME;
    Slab_Fault_History : ARRAY[0..4] OF DINT;
END_VAR
VAR
    initDone : BOOL := FALSE;
    lastValidFault : BOOL := FALSE;
    holdActive : BOOL := FALSE;
    holdElapsed : TIME := T#0MS;
    tmp_i : INT;
    tmpHoldExpired : BOOL;
    localValidFault : BOOL;
    localRising : BOOL;
END_VAR

(* ENGINEERING_CONTRACT
   THICKNESS_ALARM: active on valid-fault FALSE->TRUE (PUB001); holdActive enforces >=500ms
   using CycleTime; cleared at power-up and whenever THICKNESS_SIGNAL_VALID=FALSE (PUB004);
   remains TRUE while a valid fault persists.
   Fault record edge: logical THICKNESS_SIGNAL_VALID AND THICKNESS_FAULT false->true (PUB002).
   Counter +1, timestamp to slot 0, shift old entries 0..3 to 1..4, keep newest five.
   Runtime accumulation only when CUTTING_RUN, valid, no fault (PUB003); otherwise preserved.
   Power-up initializes all reported statistics and history to zero (PUB005).
*)

(* CONTRACT_RULES [] *)

IF NOT initDone THEN
    THICKNESS_ALARM := FALSE;
    Slab_Fault_Counter := 0;
    Slab_Runtime_Accumulator := LTIME#0S;
    FOR tmp_i := 0 TO 4 DO
        Slab_Fault_History[tmp_i] := 0;
    END_FOR;

    holdActive := FALSE;
    holdElapsed := T#0MS;
    lastValidFault := THICKNESS_SIGNAL_VALID AND THICKNESS_FAULT;
    initDone := TRUE;
    RETURN;
END_IF;

localValidFault := THICKNESS_SIGNAL_VALID AND THICKNESS_FAULT;
localRising := localValidFault AND NOT lastValidFault;

IF NOT THICKNESS_SIGNAL_VALID THEN
    THICKNESS_ALARM := FALSE;
    holdActive := FALSE;
    holdElapsed := T#0MS;
    lastValidFault := FALSE;
ELSE
    IF localRising THEN
        Slab_Fault_Counter := Slab_Fault_Counter + 1;

        FOR tmp_i := 4 TO 1 BY -1 DO
            Slab_Fault_History[tmp_i] := Slab_Fault_History[tmp_i - 1];
        END_FOR;

        Slab_Fault_History[0] := FaultTimestamp;

        holdActive := TRUE;
        holdElapsed := T#0MS;
    END_IF;

    IF holdActive THEN
        holdElapsed := holdElapsed + CycleTime;
        tmpHoldExpired := (holdElapsed >= T#500MS);
    ELSE
        tmpHoldExpired := FALSE;
    END_IF;

    THICKNESS_ALARM := localValidFault OR holdActive;

    IF tmpHoldExpired THEN
        holdActive := FALSE;
        holdElapsed := T#0MS;
    END_IF;

    IF CUTTING_RUN AND NOT THICKNESS_FAULT THEN
        Slab_Runtime_Accumulator := Slab_Runtime_Accumulator + TIME_TO_LTIME(CycleTime);
    END_IF;

    lastValidFault := localValidFault;
END_IF;
END_FUNCTION_BLOCK

(* ---- public-medium-06.candidate_02.st ---- *)
FUNCTION_BLOCK SlabThicknessFaultMonitor
VAR_INPUT
    THICKNESS_FAULT : BOOL;
    THICKNESS_SIGNAL_VALID : BOOL;
    CUTTING_RUN : BOOL;
    FaultTimestamp : DINT;
    CycleTime : TIME;
END_VAR
VAR_OUTPUT
    THICKNESS_ALARM : BOOL;
    Slab_Fault_Counter : UINT;
    Slab_Runtime_Accumulator : LTIME;
    Slab_Fault_History : ARRAY[0..4] OF DINT;
END_VAR
VAR
    initDone : BOOL := FALSE;
    lastValidFault : BOOL := FALSE;
    holdActive : BOOL := FALSE;
    holdElapsed : TIME := T#0MS;
    tmp_i : INT;
    tmpHoldExpired : BOOL;
    localValidFault : BOOL;
    localRising : BOOL;
END_VAR

(* ENGINEERING_CONTRACT
   THICKNESS_ALARM: active on valid-fault FALSE->TRUE (PUB001); holdActive enforces >=500ms
   using CycleTime; cleared at power-up and whenever THICKNESS_SIGNAL_VALID=FALSE (PUB004);
   remains TRUE while a valid fault persists.
   Fault record edge: logical THICKNESS_SIGNAL_VALID AND THICKNESS_FAULT false->true (PUB002).
   lastValidFault initialised FALSE, so first valid TRUE is a transition.
   Counter +1, timestamp to slot 0, shift old entries 0..3 to 1..4, keep newest five.
   Runtime accumulation only when CUTTING_RUN, valid, no fault (PUB003); otherwise preserved.
   Power-up initialises all reported statistics and history to zero (PUB005).
*)

(* CONTRACT_RULES [] *)

IF NOT initDone THEN
    THICKNESS_ALARM := FALSE;
    Slab_Fault_Counter := 0;
    Slab_Runtime_Accumulator := LTIME#0S;
    FOR tmp_i := 0 TO 4 DO
        Slab_Fault_History[tmp_i] := 0;
    END_FOR;

    holdActive := FALSE;
    holdElapsed := T#0MS;
    lastValidFault := FALSE;
    initDone := TRUE;
    (* No RETURN here: first invocation must also evaluate current inputs *)
END_IF;

localValidFault := THICKNESS_SIGNAL_VALID AND THICKNESS_FAULT;
localRising := localValidFault AND NOT lastValidFault;

IF NOT THICKNESS_SIGNAL_VALID THEN
    THICKNESS_ALARM := FALSE;
    holdActive := FALSE;
    holdElapsed := T#0MS;
    lastValidFault := FALSE;
ELSE
    IF localRising THEN
        Slab_Fault_Counter := Slab_Fault_Counter + 1;

        FOR tmp_i := 4 TO 1 BY -1 DO
            Slab_Fault_History[tmp_i] := Slab_Fault_History[tmp_i - 1];
        END_FOR;

        Slab_Fault_History[0] := FaultTimestamp;

        holdActive := TRUE;
        holdElapsed := T#0MS;
    END_IF;

    IF holdActive THEN
        holdElapsed := holdElapsed + CycleTime;
        tmpHoldExpired := (holdElapsed >= T#500MS);
    ELSE
        tmpHoldExpired := FALSE;
    END_IF;

    THICKNESS_ALARM := localValidFault OR holdActive;

    IF tmpHoldExpired THEN
        holdActive := FALSE;
        holdElapsed := T#0MS;
    END_IF;

    IF CUTTING_RUN AND NOT THICKNESS_FAULT THEN
        Slab_Runtime_Accumulator := Slab_Runtime_Accumulator + TIME_TO_LTIME(CycleTime);
    END_IF;

    lastValidFault := localValidFault;
END_IF;
END_FUNCTION_BLOCK

(* ---- public-medium-06.raw_candidate_01.st ---- *)
FUNCTION_BLOCK SlabThicknessFaultMonitor
VAR_INPUT
    THICKNESS_FAULT : BOOL;
    THICKNESS_SIGNAL_VALID : BOOL;
    CUTTING_RUN : BOOL;
    FaultTimestamp : DINT;
    CycleTime : TIME;
END_VAR
VAR_OUTPUT
    THICKNESS_ALARM : BOOL;
    Slab_Fault_Counter : UINT;
    Slab_Runtime_Accumulator : LTIME;
    Slab_Fault_History : ARRAY[0..4] OF DINT;
END_VAR
VAR
    initDone : BOOL := FALSE;
    lastValidFault : BOOL := FALSE;
    holdActive : BOOL := FALSE;
    holdElapsed : TIME := T#0MS;
    tmp_i : INT;
    tmpHoldExpired : BOOL;
    localValidFault : BOOL;
    localRising : BOOL;
END_VAR

(* ENGINEERING_CONTRACT
   THICKNESS_ALARM: active on valid-fault FALSE->TRUE (PUB001); holdActive enforces >=500ms
   using CycleTime; cleared at power-up and whenever THICKNESS_SIGNAL_VALID=FALSE (PUB004);
   remains TRUE while a valid fault persists.
   Fault record edge: logical THICKNESS_SIGNAL_VALID AND THICKNESS_FAULT false->true (PUB002).
   Counter +1, timestamp to slot 0, shift old entries 0..3 to 1..4, keep newest five.
   Runtime accumulation only when CUTTING_RUN, valid, no fault (PUB003); otherwise preserved.
   Power-up initializes all reported statistics and history to zero (PUB005).
*)

(* CONTRACT_RULES [] *)

IF NOT initDone THEN
    THICKNESS_ALARM := FALSE;
    Slab_Fault_Counter := 0;
    Slab_Runtime_Accumulator := LTIME#0S;
    FOR tmp_i := 0 TO 4 DO
        Slab_Fault_History[tmp_i] := 0;
    END_FOR;

    holdActive := FALSE;
    holdElapsed := T#0MS;
    lastValidFault := THICKNESS_SIGNAL_VALID AND THICKNESS_FAULT;
    initDone := TRUE;
    RETURN;
END_IF;

localValidFault := THICKNESS_SIGNAL_VALID AND THICKNESS_FAULT;
localRising := localValidFault AND NOT lastValidFault;

IF NOT THICKNESS_SIGNAL_VALID THEN
    THICKNESS_ALARM := FALSE;
    holdActive := FALSE;
    holdElapsed := T#0MS;
    lastValidFault := FALSE;
ELSE
    IF localRising THEN
        Slab_Fault_Counter := Slab_Fault_Counter + 1;

        FOR tmp_i := 4 TO 1 BY -1 DO
            Slab_Fault_History[tmp_i] := Slab_Fault_History[tmp_i - 1];
        END_FOR;

        Slab_Fault_History[0] := FaultTimestamp;

        holdActive := TRUE;
        holdElapsed := T#0MS;
    END_IF;

    IF holdActive THEN
        holdElapsed := holdElapsed + CycleTime;
        tmpHoldExpired := (holdElapsed >= T#500MS);
    ELSE
        tmpHoldExpired := FALSE;
    END_IF;

    THICKNESS_ALARM := localValidFault OR holdActive;

    IF tmpHoldExpired THEN
        holdActive := FALSE;
        holdElapsed := T#0MS;
    END_IF;

    IF CUTTING_RUN AND NOT THICKNESS_FAULT THEN
        Slab_Runtime_Accumulator := Slab_Runtime_Accumulator + TIME_TO_LTIME(CycleTime);
    END_IF;

    lastValidFault := localValidFault;
END_IF;
END_FUNCTION_BLOCK

(* ---- public-medium-06.raw_candidate_02.st ---- *)
FUNCTION_BLOCK SlabThicknessFaultMonitor
VAR_INPUT
    THICKNESS_FAULT : BOOL;
    THICKNESS_SIGNAL_VALID : BOOL;
    CUTTING_RUN : BOOL;
    FaultTimestamp : DINT;
    CycleTime : TIME;
END_VAR
VAR_OUTPUT
    THICKNESS_ALARM : BOOL;
    Slab_Fault_Counter : UINT;
    Slab_Runtime_Accumulator : LTIME;
    Slab_Fault_History : ARRAY[0..4] OF DINT;
END_VAR
VAR
    initDone : BOOL := FALSE;
    lastValidFault : BOOL := FALSE;
    holdActive : BOOL := FALSE;
    holdElapsed : TIME := T#0MS;
    tmp_i : INT;
    tmpHoldExpired : BOOL;
    localValidFault : BOOL;
    localRising : BOOL;
END_VAR

(* ENGINEERING_CONTRACT
   THICKNESS_ALARM: active on valid-fault FALSE->TRUE (PUB001); holdActive enforces >=500ms
   using CycleTime; cleared at power-up and whenever THICKNESS_SIGNAL_VALID=FALSE (PUB004);
   remains TRUE while a valid fault persists.
   Fault record edge: logical THICKNESS_SIGNAL_VALID AND THICKNESS_FAULT false->true (PUB002).
   lastValidFault initialised FALSE, so first valid TRUE is a transition.
   Counter +1, timestamp to slot 0, shift old entries 0..3 to 1..4, keep newest five.
   Runtime accumulation only when CUTTING_RUN, valid, no fault (PUB003); otherwise preserved.
   Power-up initialises all reported statistics and history to zero (PUB005).
*)

(* CONTRACT_RULES [] *)

IF NOT initDone THEN
    THICKNESS_ALARM := FALSE;
    Slab_Fault_Counter := 0;
    Slab_Runtime_Accumulator := LTIME#0S;
    FOR tmp_i := 0 TO 4 DO
        Slab_Fault_History[tmp_i] := 0;
    END_FOR;

    holdActive := FALSE;
    holdElapsed := T#0MS;
    lastValidFault := FALSE;
    initDone := TRUE;
    (* No RETURN here: first invocation must also evaluate current inputs *)
END_IF;

localValidFault := THICKNESS_SIGNAL_VALID AND THICKNESS_FAULT;
localRising := localValidFault AND NOT lastValidFault;

IF NOT THICKNESS_SIGNAL_VALID THEN
    THICKNESS_ALARM := FALSE;
    holdActive := FALSE;
    holdElapsed := T#0MS;
    lastValidFault := FALSE;
ELSE
    IF localRising THEN
        Slab_Fault_Counter := Slab_Fault_Counter + 1;

        FOR tmp_i := 4 TO 1 BY -1 DO
            Slab_Fault_History[tmp_i] := Slab_Fault_History[tmp_i - 1];
        END_FOR;

        Slab_Fault_History[0] := FaultTimestamp;

        holdActive := TRUE;
        holdElapsed := T#0MS;
    END_IF;

    IF holdActive THEN
        holdElapsed := holdElapsed + CycleTime;
        tmpHoldExpired := (holdElapsed >= T#500MS);
    ELSE
        tmpHoldExpired := FALSE;
    END_IF;

    THICKNESS_ALARM := localValidFault OR holdActive;

    IF tmpHoldExpired THEN
        holdActive := FALSE;
        holdElapsed := T#0MS;
    END_IF;

    IF CUTTING_RUN AND NOT THICKNESS_FAULT THEN
        Slab_Runtime_Accumulator := Slab_Runtime_Accumulator + TIME_TO_LTIME(CycleTime);
    END_IF;

    lastValidFault := localValidFault;
END_IF;
END_FUNCTION_BLOCK

(* ---- public-medium-07.candidate_01.st ---- *)
FUNCTION_BLOCK Office_HVAC_MultiMode_EnergySaving
VAR_INPUT
    OCCUPANCY_DETECTED : BOOL;
    ENERGY_SAVING_MODE : BOOL;
    HVAC_MODE_SELECTOR : INT;
END_VAR
VAR_OUTPUT
    SUPPLY_FAN_RUN : BOOL;
    TEMP_SETPOINT_ADJUST : INT;
END_VAR
VAR
    local_FanStart : BOOL;
    local_FanTimer : TON;
    local_TempAdjust : INT;
END_VAR

(* ENGINEERING_CONTRACT
   SUPPLY_FAN_RUN: active only after 30 s continuous OCCUPANCY_DETECTED=TRUE and Night not selected (PUB002).
   SUPPLY_FAN_RUN: reset immediately if occupancy lost or Night selected; TON resets and full 30 s required again (PUB002).
   SUPPLY_FAN_RUN: BOOL enable only; no continuous speed ramp (PUB007).
   TEMP_SETPOINT_ADJUST: combinational from current mode, occupancy and Auto-only energy-saving flag (PUB003/PUB004/PUB005).
   TEMP_SETPOINT_ADJUST: INT degrees C, clamped to [-4,4]; no retention or explicit reset (PUB006).
   Initialization: variables start FALSE/0; normal calculation then updates outputs from current inputs (PUB006).
   Valid selector values are 0..3; callers guarantee this (PUB001). Invalid selector handling is unspecified and maps to 0 C adjustment.
*)

(* CONTRACT_RULES [] *)

local_FanStart := OCCUPANCY_DETECTED AND (HVAC_MODE_SELECTOR <> 3);

local_FanTimer(IN := local_FanStart, PT := T#30S);
SUPPLY_FAN_RUN := local_FanTimer.Q;

CASE HVAC_MODE_SELECTOR OF
    0: (* Auto *)
        IF OCCUPANCY_DETECTED THEN
            local_TempAdjust := 0;
        ELSIF ENERGY_SAVING_MODE THEN
            local_TempAdjust := 3;
        ELSE
            local_TempAdjust := 2;
        END_IF;

    1: (* Comfort *)
        IF OCCUPANCY_DETECTED THEN
            local_TempAdjust := 0;
        ELSE
            local_TempAdjust := 1;
        END_IF;

    2: (* Economy *)
        IF OCCUPANCY_DETECTED THEN
            local_TempAdjust := 0;
        ELSE
            local_TempAdjust := 4;
        END_IF;

    3: (* Night *)
        local_TempAdjust := 4;

ELSE
    local_TempAdjust := 0; (* unspecified invalid input handling *)
END_CASE;

IF local_TempAdjust > 4 THEN
    local_TempAdjust := 4;
ELSIF local_TempAdjust < -4 THEN
    local_TempAdjust := -4;
END_IF;

TEMP_SETPOINT_ADJUST := local_TempAdjust;

END_FUNCTION_BLOCK

(* ---- public-medium-07.raw_candidate_01.st ---- *)
FUNCTION_BLOCK Office_HVAC_MultiMode_EnergySaving
VAR_INPUT
    OCCUPANCY_DETECTED : BOOL;
    ENERGY_SAVING_MODE : BOOL;
    HVAC_MODE_SELECTOR : INT;
END_VAR
VAR_OUTPUT
    SUPPLY_FAN_RUN : BOOL;
    TEMP_SETPOINT_ADJUST : INT;
END_VAR
VAR
    local_FanStart : BOOL;
    local_FanTimer : TON;
    local_TempAdjust : INT;
END_VAR

(* ENGINEERING_CONTRACT
   SUPPLY_FAN_RUN: active only after 30 s continuous OCCUPANCY_DETECTED=TRUE and Night not selected (PUB002).
   SUPPLY_FAN_RUN: reset immediately if occupancy lost or Night selected; TON resets and full 30 s required again (PUB002).
   SUPPLY_FAN_RUN: BOOL enable only; no continuous speed ramp (PUB007).
   TEMP_SETPOINT_ADJUST: combinational from current mode, occupancy and Auto-only energy-saving flag (PUB003/PUB004/PUB005).
   TEMP_SETPOINT_ADJUST: INT degrees C, clamped to [-4,4]; no retention or explicit reset (PUB006).
   Initialization: variables start FALSE/0; normal calculation then updates outputs from current inputs (PUB006).
   Valid selector values are 0..3; callers guarantee this (PUB001). Invalid selector handling is unspecified and maps to 0 C adjustment.
*)

(* CONTRACT_RULES [] *)

local_FanStart := OCCUPANCY_DETECTED AND (HVAC_MODE_SELECTOR <> 3);

local_FanTimer(IN := local_FanStart, PT := T#30S);
SUPPLY_FAN_RUN := local_FanTimer.Q;

CASE HVAC_MODE_SELECTOR OF
    0: (* Auto *)
        IF OCCUPANCY_DETECTED THEN
            local_TempAdjust := 0;
        ELSIF ENERGY_SAVING_MODE THEN
            local_TempAdjust := 3;
        ELSE
            local_TempAdjust := 2;
        END_IF;

    1: (* Comfort *)
        IF OCCUPANCY_DETECTED THEN
            local_TempAdjust := 0;
        ELSE
            local_TempAdjust := 1;
        END_IF;

    2: (* Economy *)
        IF OCCUPANCY_DETECTED THEN
            local_TempAdjust := 0;
        ELSE
            local_TempAdjust := 4;
        END_IF;

    3: (* Night *)
        local_TempAdjust := 4;

ELSE
    local_TempAdjust := 0; (* unspecified invalid input handling *)
END_CASE;

IF local_TempAdjust > 4 THEN
    local_TempAdjust := 4;
ELSIF local_TempAdjust < -4 THEN
    local_TempAdjust := -4;
END_IF;

TEMP_SETPOINT_ADJUST := local_TempAdjust;

END_FUNCTION_BLOCK

(* ---- public-medium-08.candidate_01.st ---- *)
(*
ENGINEERING_CONTRACT
ipValue: combinational UDINT, set every invocation to parsed IPv4 in network byte order (PUB002).
Invalid/malformed input, nondigit, wrong segment count, or octet >255 forces ipValue := 0 (PUB003).
No retention, no latch, no reset; each scan recomputes independently.
Same-scan priority: partial octet shifts are discarded if any later failure occurs.
Units: octets are 0..255, 8-bit; first text segment maps to bits 31..24, last to 7..0.
Leading zeros are accepted because PUB001 forbids only non-digit/empty and enforces value range.
*)
(* CONTRACT_RULES [] *)
FUNCTION_BLOCK IPv4Parser
VAR_INPUT
    ipText : STRING(254);
END_VAR
VAR_OUTPUT
    ipValue : UDINT;
END_VAR
VAR
    tmp_len : INT;
    tmp_idx : INT;
    tmp_segCount : INT;      (* 1..4, current segment being parsed *)
    tmp_segVal : UDINT;      (* accumulated value of current segment *)
    tmp_segHasDigit : BOOL;  (* TRUE if current segment contains at least one digit *)
    tmp_parseOk : BOOL;      (* FALSE after any malformed condition *)
    tmp_char : INT;          (* ASCII code of current character *)
    tmp_digit : UDINT;       (* numeric value of current digit *)
END_VAR

ipValue := 0;
tmp_len := LEN(ipText);
tmp_idx := 0;
tmp_segCount := 1;
tmp_segVal := 0;
tmp_segHasDigit := FALSE;
tmp_parseOk := TRUE;

WHILE (tmp_idx < tmp_len) DO
    tmp_char := BYTE_TO_INT(ipText[tmp_idx]);

    IF (tmp_char >= 48) AND (tmp_char <= 57) THEN
        tmp_segHasDigit := TRUE;
        tmp_digit := INT_TO_UDINT(tmp_char - 48);
        tmp_segVal := tmp_segVal * TO_UDINT(10) + tmp_digit;

        IF tmp_segVal > 255 THEN
            tmp_parseOk := FALSE;
            EXIT;
        END_IF;

    ELSIF tmp_char = 46 THEN
        (* Dot: finalize current segment and advance to next *)
        IF (NOT tmp_segHasDigit) OR (tmp_segCount >= 4) THEN
            tmp_parseOk := FALSE;
            EXIT;
        END_IF;

        ipValue := SHL(ipValue, 8);
        ipValue := ipValue OR tmp_segVal;

        tmp_segCount := tmp_segCount + 1;
        tmp_segVal := 0;
        tmp_segHasDigit := FALSE;

    ELSE
        tmp_parseOk := FALSE;
        EXIT;
    END_IF;

    tmp_idx := tmp_idx + 1;
END_WHILE;

IF tmp_parseOk THEN
    IF (tmp_segCount <> 4) OR (NOT tmp_segHasDigit) THEN
        tmp_parseOk := FALSE;
    ELSE
        ipValue := SHL(ipValue, 8);
        ipValue := ipValue OR tmp_segVal;
    END_IF;
END_IF;

IF NOT tmp_parseOk THEN
    ipValue := 0;
END_IF;

END_FUNCTION_BLOCK

(* ---- public-medium-08.raw_candidate_01.st ---- *)
(*
ENGINEERING_CONTRACT
ipValue: combinational UDINT, set every invocation to parsed IPv4 in network byte order (PUB002).
Invalid/malformed input, nondigit, wrong segment count, or octet >255 forces ipValue := 0 (PUB003).
No retention, no latch, no reset; each scan recomputes independently.
Same-scan priority: partial octet shifts are discarded if any later failure occurs.
Units: octets are 0..255, 8-bit; first text segment maps to bits 31..24, last to 7..0.
Leading zeros are accepted because PUB001 forbids only non-digit/empty and enforces value range.
*)
(* CONTRACT_RULES [] *)
FUNCTION_BLOCK IPv4Parser
VAR_INPUT
    ipText : STRING(254);
END_VAR
VAR_OUTPUT
    ipValue : UDINT;
END_VAR
VAR
    tmp_len : INT;
    tmp_idx : INT;
    tmp_segCount : INT;      (* 1..4, current segment being parsed *)
    tmp_segVal : UDINT;      (* accumulated value of current segment *)
    tmp_segHasDigit : BOOL;  (* TRUE if current segment contains at least one digit *)
    tmp_parseOk : BOOL;      (* FALSE after any malformed condition *)
    tmp_char : INT;          (* ASCII code of current character *)
    tmp_digit : UDINT;       (* numeric value of current digit *)
END_VAR

ipValue := 0;
tmp_len := LEN(ipText);
tmp_idx := 0;
tmp_segCount := 1;
tmp_segVal := 0;
tmp_segHasDigit := FALSE;
tmp_parseOk := TRUE;

WHILE (tmp_idx < tmp_len) DO
    tmp_char := BYTE_TO_INT(ipText[tmp_idx]);

    IF (tmp_char >= 48) AND (tmp_char <= 57) THEN
        tmp_segHasDigit := TRUE;
        tmp_digit := INT_TO_UDINT(tmp_char - 48);
        tmp_segVal := tmp_segVal * TO_UDINT(10) + tmp_digit;

        IF tmp_segVal > 255 THEN
            tmp_parseOk := FALSE;
            EXIT;
        END_IF

    ELSIF tmp_char = 46 THEN
        (* Dot: finalize current segment and advance to next *)
        IF (NOT tmp_segHasDigit) OR (tmp_segCount >= 4) THEN
            tmp_parseOk := FALSE;
            EXIT;
        END_IF

        ipValue := SHL(ipValue, 8);
        ipValue := ipValue OR tmp_segVal;

        tmp_segCount := tmp_segCount + 1;
        tmp_segVal := 0;
        tmp_segHasDigit := FALSE;

    ELSE
        tmp_parseOk := FALSE;
        EXIT;
    END_IF

    tmp_idx := tmp_idx + 1;
END_WHILE

IF tmp_parseOk THEN
    IF (tmp_segCount <> 4) OR (NOT tmp_segHasDigit) THEN
        tmp_parseOk := FALSE;
    ELSE
        ipValue := SHL(ipValue, 8);
        ipValue := ipValue OR tmp_segVal;
    END_IF
END_IF

IF NOT tmp_parseOk THEN
    ipValue := 0;
END_IF

END_FUNCTION_BLOCK

(* ---- self-easy-01.candidate_01.st ---- *)
(*
ENGINEERING_CONTRACT
avgOut REAL output:
- Activation: enable AND avgEnable AND count>=1 -> avgOut = sum(values[1..min(count,8)]) / min(count,8) using DINT accumulation and REAL division.
- Hold/retention: enable=FALSE or avgEnable=FALSE or count<=0 -> avgOut := tmp_heldOut (previous value); no arithmetic or division in same scan.
- Reset/deactivation: no dedicated reset input; held value persists in VAR tmp_heldOut. Initial avgOut/tmp_heldOut = 0.0 (unspecified).
- Same-scan priority: any hold condition suppresses update; count>8 is clipped to 8 before summing.
- Units/bounds: INT samples converted to DINT; sum range max +/-262144; REAL result, no rounding; count negative not used.
*)
(* CONTRACT_RULES [] *)
FUNCTION_BLOCK FB
VAR_INPUT
    enable : BOOL;
    values : ARRAY[1..8] OF INT;
    count : INT;
    avgEnable : BOOL;
END_VAR
VAR_OUTPUT
    avgOut : REAL;
END_VAR
VAR
    tmp_sum : DINT;
    tmp_count : INT;
    tmp_i : INT;
    tmp_heldOut : REAL;
END_VAR

IF enable AND avgEnable AND (count >= 1) THEN
    IF count > 8 THEN
        tmp_count := 8;
    ELSE
        tmp_count := count;
    END_IF;

    tmp_sum := 0;
    FOR tmp_i := 1 TO tmp_count BY 1 DO
        tmp_sum := tmp_sum + INT_TO_DINT(values[tmp_i]);
    END_FOR;

    tmp_heldOut := DINT_TO_REAL(tmp_sum) / INT_TO_REAL(tmp_count);
    avgOut := tmp_heldOut;
ELSE
    avgOut := tmp_heldOut;
END_IF;

END_FUNCTION_BLOCK

(* ---- self-easy-01.raw_candidate_01.st ---- *)
(*
ENGINEERING_CONTRACT
avgOut REAL output:
- Activation: enable AND avgEnable AND count>=1 -> avgOut = sum(values[1..min(count,8)]) / min(count,8) using DINT accumulation and REAL division.
- Hold/retention: enable=FALSE or avgEnable=FALSE or count<=0 -> avgOut := tmp_heldOut (previous value); no arithmetic or division in same scan.
- Reset/deactivation: no dedicated reset input; held value persists in VAR tmp_heldOut. Initial avgOut/tmp_heldOut = 0.0 (unspecified).
- Same-scan priority: any hold condition suppresses update; count>8 is clipped to 8 before summing.
- Units/bounds: INT samples converted to DINT; sum range max +/-262144; REAL result, no rounding; count negative not used.
*)
(* CONTRACT_RULES [] *)
FUNCTION_BLOCK FB
VAR_INPUT
    enable : BOOL;
    values : ARRAY[1..8] OF INT;
    count : INT;
    avgEnable : BOOL;
END_VAR
VAR_OUTPUT
    avgOut : REAL;
END_VAR
VAR
    tmp_sum : DINT;
    tmp_count : INT;
    tmp_i : INT;
    tmp_heldOut : REAL;
END_VAR

IF enable AND avgEnable AND (count >= 1) THEN
    IF count > 8 THEN
        tmp_count := 8;
    ELSE
        tmp_count := count;
    END_IF;

    tmp_sum := 0;
    FOR tmp_i := 1 TO tmp_count BY 1 DO
        tmp_sum := tmp_sum + INT_TO_DINT(values[tmp_i]);
    END_FOR;

    tmp_heldOut := DINT_TO_REAL(tmp_sum) / INT_TO_REAL(tmp_count);
    avgOut := tmp_heldOut;
ELSE
    avgOut := tmp_heldOut;
END_IF;

END_FUNCTION_BLOCK

(* ---- self-easy-02.candidate_01.st ---- *)
(* ENGINEERING_CONTRACT
   alarmHigh: set when tankLevel >= 85.0; latch until rising resetBtn while high danger absent.
   alarmLow:  set when tankLevel <= 15.0; latch until rising resetBtn while low danger absent.
   Danger has same-scan priority over reset.
   reset edge = resetBtn AND NOT prevResetBtn; prevResetBtn initial FALSE.
   pumpRun = inletPermit AND NOT alarmHigh AND NOT alarmLow after alarm update.
   outletValveOpen = NOT alarmLow.
   outletFlow is unused in this function block.
   All outputs sampled at end of the same scan.
*)
(* CONTRACT_RULES [] *)
FUNCTION_BLOCK FB
VAR_INPUT
    tankLevel : REAL;
    outletFlow : REAL;
    inletPermit : BOOL;
    resetBtn : BOOL;
END_VAR
VAR_OUTPUT
    pumpRun : BOOL;
    alarmHigh : BOOL;
    alarmLow : BOOL;
    outletValveOpen : BOOL;
END_VAR
VAR
    prevResetBtn : BOOL := FALSE;
    prevAlarmHigh : BOOL := FALSE;
    prevAlarmLow : BOOL := FALSE;
    tmp_highDanger : BOOL;
    tmp_lowDanger : BOOL;
    tmp_resetEdge : BOOL;
    tmp_newHigh : BOOL;
    tmp_newLow : BOOL;
END_VAR

tmp_highDanger := tankLevel >= 85.0;
tmp_lowDanger := tankLevel <= 15.0;
tmp_resetEdge := resetBtn AND NOT prevResetBtn;

IF tmp_highDanger THEN
    tmp_newHigh := TRUE;
ELSIF tmp_resetEdge THEN
    tmp_newHigh := FALSE;
ELSE
    tmp_newHigh := prevAlarmHigh;
END_IF;

IF tmp_lowDanger THEN
    tmp_newLow := TRUE;
ELSIF tmp_resetEdge THEN
    tmp_newLow := FALSE;
ELSE
    tmp_newLow := prevAlarmLow;
END_IF;

alarmHigh := tmp_newHigh;
alarmLow := tmp_newLow;

pumpRun := inletPermit AND NOT alarmHigh AND NOT alarmLow;
outletValveOpen := NOT alarmLow;

prevResetBtn := resetBtn;
prevAlarmHigh := alarmHigh;
prevAlarmLow := alarmLow;

END_FUNCTION_BLOCK

(* ---- self-easy-02.raw_candidate_01.st ---- *)
(* ENGINEERING_CONTRACT
   alarmHigh: set when tankLevel >= 85.0; latch until rising resetBtn while high danger absent.
   alarmLow:  set when tankLevel <= 15.0; latch until rising resetBtn while low danger absent.
   Danger has same-scan priority over reset.
   reset edge = resetBtn AND NOT prevResetBtn; prevResetBtn initial FALSE.
   pumpRun = inletPermit AND NOT alarmHigh AND NOT alarmLow after alarm update.
   outletValveOpen = NOT alarmLow.
   outletFlow is unused in this function block.
   All outputs sampled at end of the same scan.
*)
(* CONTRACT_RULES [] *)
FUNCTION_BLOCK FB
VAR_INPUT
    tankLevel : REAL;
    outletFlow : REAL;
    inletPermit : BOOL;
    resetBtn : BOOL;
END_VAR
VAR_OUTPUT
    pumpRun : BOOL;
    alarmHigh : BOOL;
    alarmLow : BOOL;
    outletValveOpen : BOOL;
END_VAR
VAR
    prevResetBtn : BOOL := FALSE;
    prevAlarmHigh : BOOL := FALSE;
    prevAlarmLow : BOOL := FALSE;
    tmp_highDanger : BOOL;
    tmp_lowDanger : BOOL;
    tmp_resetEdge : BOOL;
    tmp_newHigh : BOOL;
    tmp_newLow : BOOL;
END_VAR

tmp_highDanger := tankLevel >= 85.0;
tmp_lowDanger := tankLevel <= 15.0;
tmp_resetEdge := resetBtn AND NOT prevResetBtn;

IF tmp_highDanger THEN
    tmp_newHigh := TRUE;
ELSIF tmp_resetEdge THEN
    tmp_newHigh := FALSE;
ELSE
    tmp_newHigh := prevAlarmHigh;
END_IF;

IF tmp_lowDanger THEN
    tmp_newLow := TRUE;
ELSIF tmp_resetEdge THEN
    tmp_newLow := FALSE;
ELSE
    tmp_newLow := prevAlarmLow;
END_IF;

alarmHigh := tmp_newHigh;
alarmLow := tmp_newLow;

pumpRun := inletPermit AND NOT alarmHigh AND NOT alarmLow;
outletValveOpen := NOT alarmLow;

prevResetBtn := resetBtn;
prevAlarmHigh := alarmHigh;
prevAlarmLow := alarmLow;

END_FUNCTION_BLOCK

(* ---- self-hard-01.candidate_01.st ---- *)
FUNCTION_BLOCK FB
VAR_INPUT
    flowLow: BOOL;
    ackBtn: BOOL;
    sensorOK: BOOL;
END_VAR
VAR_OUTPUT
    alarmActive: BOOL;
    alarmAcked: BOOL;
    highHigh: BOOL;
END_VAR
VAR
    prev_flowLow: BOOL := FALSE;
    prev_ackBtn: BOOL := FALSE;
    prev_alarmActive: BOOL := FALSE;
    prev_alarmAcked: BOOL := FALSE;
    rising_ack: BOOL;
    prev_combined: BOOL;
    prev_triple: BOOL;
    new_alarmActive: BOOL;
    new_alarmAcked: BOOL;
END_VAR

(* ENGINEERING_CONTRACT
   alarmActive: state latch; activates on flowLow TRUE (PUB001-PUB003);
     retains while prior alarmActive TRUE and no ack rising edge and not
     prior (flowLow AND alarmAcked); clears only on ack rising edge when
     flowLow FALSE (PUB003, S6). Same-scan independent of highHigh.
   alarmAcked: state latch; set when alarmActive and either flowLow FALSE,
     ack rising edge, or prior (flowLow AND alarmActive AND alarmAcked);
     clears with alarmActive (PUB002-PUB003, S7).
   highHigh: pure combinational; TRUE exactly when sensorOK FALSE;
     no retention; same-scan (PUB004-PUB005, S3, S5).
   All states updated once per scan; outputs sampled at cycle end.
*)

(* CONTRACT_RULES [] *)

highHigh := NOT sensorOK;

rising_ack := ackBtn AND NOT prev_ackBtn;

prev_combined := prev_flowLow AND prev_alarmAcked;
prev_triple := prev_flowLow AND prev_alarmActive AND prev_alarmAcked;

new_alarmActive := flowLow OR (prev_alarmActive AND NOT rising_ack AND NOT prev_combined);
new_alarmAcked := new_alarmActive AND (NOT flowLow OR rising_ack OR prev_triple);

alarmActive := new_alarmActive;
alarmAcked := new_alarmAcked;

prev_flowLow := flowLow;
prev_ackBtn := ackBtn;
prev_alarmActive := alarmActive;
prev_alarmAcked := alarmAcked;

END_FUNCTION_BLOCK

(* ---- self-hard-01.raw_candidate_01.st ---- *)
FUNCTION_BLOCK FB
VAR_INPUT
    flowLow: BOOL;
    ackBtn: BOOL;
    sensorOK: BOOL;
END_VAR
VAR_OUTPUT
    alarmActive: BOOL;
    alarmAcked: BOOL;
    highHigh: BOOL;
END_VAR
VAR
    prev_flowLow: BOOL := FALSE;
    prev_ackBtn: BOOL := FALSE;
    prev_alarmActive: BOOL := FALSE;
    prev_alarmAcked: BOOL := FALSE;
    rising_ack: BOOL;
    prev_combined: BOOL;
    prev_triple: BOOL;
    new_alarmActive: BOOL;
    new_alarmAcked: BOOL;
END_VAR

(* ENGINEERING_CONTRACT
   alarmActive: state latch; activates on flowLow TRUE (PUB001-PUB003);
     retains while prior alarmActive TRUE and no ack rising edge and not
     prior (flowLow AND alarmAcked); clears only on ack rising edge when
     flowLow FALSE (PUB003, S6). Same-scan independent of highHigh.
   alarmAcked: state latch; set when alarmActive and either flowLow FALSE,
     ack rising edge, or prior (flowLow AND alarmActive AND alarmAcked);
     clears with alarmActive (PUB002-PUB003, S7).
   highHigh: pure combinational; TRUE exactly when sensorOK FALSE;
     no retention; same-scan (PUB004-PUB005, S3, S5).
   All states updated once per scan; outputs sampled at cycle end.
*)

(* CONTRACT_RULES [] *)

highHigh := NOT sensorOK;

rising_ack := ackBtn AND NOT prev_ackBtn;

prev_combined := prev_flowLow AND prev_alarmAcked;
prev_triple := prev_flowLow AND prev_alarmActive AND prev_alarmAcked;

new_alarmActive := flowLow OR (prev_alarmActive AND NOT rising_ack AND NOT prev_combined);
new_alarmAcked := new_alarmActive AND (NOT flowLow OR rising_ack OR prev_triple);

alarmActive := new_alarmActive;
alarmAcked := new_alarmAcked;

prev_flowLow := flowLow;
prev_ackBtn := ackBtn;
prev_alarmActive := alarmActive;
prev_alarmAcked := alarmAcked;

END_FUNCTION_BLOCK

(* ---- self-hard-02.candidate_01.st ---- *)
(* ENGINEERING_CONTRACT
   - phase: 0 idle initial; new start & !abort -> 1; in running, elapsed<maxDuration and (prevPhase=2 or pv>=setpoint) -> 2, else 1; elapsed>=maxDuration -> 3; abort -> 9. Priority abort > start edge > run count (PUB002-006).
   - elapsed: increment exactly once per scan when !abort, !startEdge, prevPhase=1/2; reset 0 on new start; freeze otherwise.
   - timeout: set TRUE exactly when running scan counted reaches maxDuration; reset FALSE on new start; freeze on abort/completion/idle.
   - start rising edge recorded first and consumed even if abort same scan; restart requires release/press.
   - maxDuration positive scan count; comparison >=. Boundaries: counts scan after start not counted.
*)
FUNCTION_BLOCK FB
VAR
    prevStartBtn : BOOL := FALSE;
    prevPhase : INT := 0;
    prevElapsed : INT := 0;
    prevTimeout : BOOL := FALSE;
    startEdge : BOOL;
END_VAR

(* Record startBtn rising edge before priority processing; consumed even if abort *)
startEdge := startBtn AND NOT prevStartBtn;

IF abortBtn THEN
    (* Abort has highest priority: enter phase 9 and freeze elapsed/timeout *)
    phase := 9;
    elapsed := prevElapsed;
    timeout := prevTimeout;
ELSIF startEdge THEN
    (* New valid start with no abort: reset batch and do not count this scan *)
    phase := 1;
    elapsed := 0;
    timeout := FALSE;
ELSE
    (* No abort and no new start edge *)
    IF (prevPhase = 1) OR (prevPhase = 2) THEN
        (* Running state: count exactly one scan *)
        elapsed := prevElapsed + 1;

        IF elapsed >= maxDuration THEN
            (* Timeout has priority over temperature threshold *)
            timeout := TRUE;
            phase := 3;
        ELSE
            timeout := FALSE;
            IF (prevPhase = 2) OR (pv >= setpoint) THEN
                phase := 2;
            ELSE
                phase := 1;
            END_IF;
        END_IF;
    ELSE
        (* Idle, complete, or aborted: hold state *)
        phase := prevPhase;
        elapsed := prevElapsed;
        timeout := prevTimeout;
    END_IF;
END_IF;

(* Update previous-cycle memory *)
prevStartBtn := startBtn;
prevPhase := phase;
prevElapsed := elapsed;
prevTimeout := timeout;

(* CONTRACT_RULES [] *)
END_FUNCTION_BLOCK
